FBuilder.Initialize(Mode := E_OrchestrationMode.ParallelSlots,
    TestCases := FCases);
AcceptedA := FBuilder.RegisterWithSlot(TestCase := ChildA,
    ExecutionSlot := 0);
Config := FBuilder.Finalize();
FZeroSlotRejectedMatches := NOT AcceptedA AND NOT Config.IsValid
    AND (FBuilder.Count = 0) AND (FCases[1] = 0)
    AND (FChildA.ExecutionSlot = CandidateSlotBeforeRejection);

FBuilder.Initialize(Mode := E_OrchestrationMode.ParallelSlots,
    TestCases := FCases);
AcceptedA := FBuilder.RegisterWithSlot(TestCase := ChildA,
    ExecutionSlot := 1);
AcceptedB := FBuilder.RegisterWithSlot(TestCase := ChildB,
    ExecutionSlot := 3);
Config := FBuilder.Finalize();
FSlotGapRejectedMatches := AcceptedA AND AcceptedB AND NOT Config.IsValid
    AND FBuilder.IsFinalized AND (FBuilder.Count = 2)
    AND (FCases[1] = ChildA) AND (FCases[2] = ChildB);
END_METHOD

END_FUNCTION_BLOCK

// ---- SelfTests/TestCases/TestSuite_TestSuiteConfigurationBuilder/Test_SuiteBuilderFinalizeReuse.TcPOU
{region 'Documentation'}
(*!
<summary>Checks empty and repeated finalization, sealed registration and a clean new build.</summary>
<description>Child mocks are inert interface identities and slot storage only; no child initialization or FB call is performed.</description>
*)
{endregion}
FUNCTION_BLOCK Test_SuiteBuilderFinalizeReuse EXTENDS TestCaseBase
VAR
    FBuilder : TestSuiteConfigurationBuilder;
    FCases : ARRAY[1..2] OF I_TestCase;
    FChildA : TestCaseMock;
    FChildB : TestCaseMock;
    FScenarioExecuted : BOOL;
    FChecksEvaluated : BOOL;
    FEmptyRejected : AssertTrue;
    FEmptyRejectedMatches : BOOL;
    FRepeatedFinalization : AssertTrue;
    FRepeatedFinalizationMatches : BOOL;
    FSealedRegistration : AssertTrue;
    FSealedRegistrationMatches : BOOL;
    FErrorRecorded : AssertTrue;
    FErrorRecordedMatches : BOOL;
    FFreshInitialize : AssertTrue;
    FFreshInitializeMatches : BOOL;
    FReuse : AssertTrue;
    FReuseMatches : BOOL;
END_VAR
VAR CONSTANT
    CandidateSlotBeforeRejection : UINT := 9;
END_VAR

SUPER^();

{region 'Documentation'}
(*!
<summary>Contributes each owned Assertion once without executing it.</summary>
*)
{endregion}
METHOD PROTECTED AggregateResults
VAR_INPUT
    Aggregator : I_ResultAggregator; //! Borrowed result sink owned by the outer Test Case; add this test's checking Assertions without resetting or retaining the sink.
END_VAR
Aggregator.AddProvider(Provider := FEmptyRejected);
Aggregator.AddProvider(Provider := FRepeatedFinalization);
Aggregator.AddProvider(Provider := FSealedRegistration);
Aggregator.AddProvider(Provider := FErrorRecorded);
Aggregator.AddProvider(Provider := FFreshInitialize);
Aggregator.AddProvider(Provider := FReuse);
END_METHOD

{region 'Documentation'}
(*!
<summary>Requires successful base and owned Assertion initialization.</summary>
*)
{endregion}
METHOD PROTECTED CheckInitialization : BOOL //! TRUE when the inherited initialization check and this concrete fixture check both accept the setup.
CheckInitialization := FALSE;
IF NOT SUPER^.CheckInitialization() THEN
    RETURN;
END_IF;

CheckInitialization := FEmptyRejected.IsInitialized
    AND FRepeatedFinalization.IsInitialized
    AND FSealedRegistration.IsInitialized
    AND FErrorRecorded.IsInitialized
    AND FFreshInitialize.IsInitialized
    AND FReuse.IsInitialized;
END_METHOD

{region 'Documentation'}
(*!
<summary>Configures one direct builder scenario and its named Assertions.</summary>
*)
{endregion}
METHOD PROTECTED Configure
FPreparationStateCount := 0;
FTestStateCount := 1;
FScenarioExecuted := FALSE;
FChecksEvaluated := FALSE;

FEmptyRejectedMatches := FALSE;
FEmptyRejected.Initialize(Parent := THIS^,
    AssertionName := 'EmptyRejected');
FRepeatedFinalizationMatches := FALSE;
FRepeatedFinalization.Initialize(Parent := THIS^,
    AssertionName := 'RepeatedFinalization');
FSealedRegistrationMatches := FALSE;
FSealedRegistration.Initialize(Parent := THIS^,
    AssertionName := 'SealedRegistration');
FErrorRecordedMatches := FALSE;
FErrorRecorded.Initialize(Parent := THIS^,
    AssertionName := 'ErrorRecorded');
FFreshInitializeMatches := FALSE;
FFreshInitialize.Initialize(Parent := THIS^,
    AssertionName := 'FreshInitialize');
FReuseMatches := FALSE;
FReuse.Initialize(Parent := THIS^,
    AssertionName := 'Reuse');
END_METHOD

{region 'Documentation'}
(*!
<summary>Completes Abort immediately; no asynchronous resource operation is started.</summary>
*)
{endregion}
METHOD PROTECTED ProcessAbort
VAR_INPUT
    Enable : BOOL; //! Phase permission supplied by the owning Test Case; FALSE does not authorize progression, while observation may continue.
END_VAR
IF Enable THEN
    CompleteAbort();
END_IF;
END_METHOD

{region 'Documentation'}
(*!
<summary>Evaluates recorded observations and consumes pending resets on disabled calls.</summary>
*)
{endregion}
METHOD PROTECTED ProcessAssertions
VAR_INPUT
    Enable : BOOL; //! Phase permission supplied by the owning Test Case; FALSE does not authorize progression, while observation may continue.
END_VAR
FEmptyRejected(Enable := Enable,
    State := State,
    IN := FEmptyRejectedMatches);

FRepeatedFinalization(Enable := Enable,
    State := State,
    IN := FRepeatedFinalizationMatches);

FSealedRegistration(Enable := Enable,
    State := State,
    IN := FSealedRegistrationMatches);

FErrorRecorded(Enable := Enable,
    State := State,
    IN := FErrorRecordedMatches);

FFreshInitialize(Enable := Enable,
    State := State,
    IN := FFreshInitializeMatches);

FReuse(Enable := Enable,
    State := State,
    IN := FReuseMatches);

IF Enable AND FEmptyRejected.EvaluationActive
    AND FRepeatedFinalization.EvaluationActive
    AND FSealedRegistration.EvaluationActive
    AND FErrorRecorded.EvaluationActive
    AND FFreshInitialize.EvaluationActive
    AND FReuse.EvaluationActive THEN
    FChecksEvaluated := TRUE;
END_IF;
END_METHOD

{region 'Documentation'}
(*!
<summary>No Preparation phase is needed for synchronous builder calls.</summary>
*)
{endregion}
METHOD PROTECTED ProcessPreparations
VAR_INPUT
    // SA0033: Required override signature; this scenario has no Preparation work.
    {attribute 'analysis' := '-33'}
    Enable : BOOL; //! Phase permission supplied by the owning Test Case; FALSE does not authorize progression, while observation may continue.
END_VAR
END_METHOD

{region 'Documentation'}
(*!
<summary>Clears recorded checks and Assertion results; each scenario initializes its own builder.</summary>
*)
{endregion}
METHOD PROTECTED ProcessReset
FScenarioExecuted := FALSE;
FChecksEvaluated := FALSE;
FEmptyRejectedMatches := FALSE;
FEmptyRejected.Reset();
FRepeatedFinalizationMatches := FALSE;
FRepeatedFinalization.Reset();
FSealedRegistrationMatches := FALSE;
FSealedRegistration.Reset();
FErrorRecordedMatches := FALSE;
FErrorRecorded.Reset();
FFreshInitializeMatches := FALSE;
FFreshInitialize.Reset();
FReuseMatches := FALSE;
FReuse.Reset();
CompleteReset();
END_METHOD

{region 'Documentation'}
(*!
<summary>Runs setup operations once, then completes after their observations have been evaluated.</summary>
*)
{endregion}
METHOD PROTECTED ProcessTests
VAR_INPUT
    Enable : BOOL; //! Phase permission supplied by the owning Test Case; FALSE does not authorize progression, while observation may continue.
END_VAR
IF NOT Enable THEN
    RETURN;
END_IF;

IF FChecksEvaluated THEN
    CompleteTests();
ELSIF NOT FScenarioExecuted THEN
    RunScenario();
    FScenarioExecuted := TRUE;
END_IF;
END_METHOD

{region 'Documentation'}
(*!
<summary>Checks empty and repeated finalization, sealed registration and a clean new build.</summary>
*)
{endregion}
METHOD PRIVATE RunScenario
VAR
    ChildA : I_TestCase;
    ChildB : I_TestCase;
    AcceptedA : BOOL;
    AcceptedB : BOOL;
    Config : ST_TestCaseCollectionConfig;
    RepeatedConfig : ST_TestCaseCollectionConfig;
END_VAR
ChildA := FChildA;
ChildB := FChildB;
FBuilder.Initialize(Mode := E_OrchestrationMode.Serial,
    TestCases := FCases);
Config := FBuilder.Finalize();
RepeatedConfig := FBuilder.Finalize();
FEmptyRejectedMatches := NOT Config.IsValid AND NOT RepeatedConfig.IsValid
    AND FBuilder.IsFinalized AND NOT FBuilder.IsValid AND (RepeatedConfig.Count = 0);

FBuilder.Initialize(Mode := E_OrchestrationMode.Serial,
    TestCases := FCases);
AcceptedA := FBuilder.Register(TestCase := ChildA);
Config := FBuilder.Finalize();
RepeatedConfig := FBuilder.Finalize();
FRepeatedFinalizationMatches := AcceptedA AND Config.IsValid AND RepeatedConfig.IsValid
    AND (RepeatedConfig.FirstIndex = Config.FirstIndex)
    AND (RepeatedConfig.LastIndex = Config.LastIndex)
    AND (RepeatedConfig.Count = Config.Count) AND (RepeatedConfig.Mode = Config.Mode);

FChildB.ExecutionSlot := CandidateSlotBeforeRejection;
AcceptedB := FBuilder.Register(TestCase := ChildB);
RepeatedConfig := FBuilder.Finalize();
FSealedRegistrationMatches := NOT AcceptedB AND RepeatedConfig.IsValid AND FBuilder.IsValid
    AND FBuilder.IsFinalized AND (FBuilder.Count = 1)
    AND (FCases[1] = ChildA) AND (FCases[2] = 0)
    AND (FChildB.ExecutionSlot = CandidateSlotBeforeRejection);

FBuilder.Initialize(Mode := E_OrchestrationMode.Serial,
    TestCases := FCases);
AcceptedA := FBuilder.Register(TestCase := ChildA);
AcceptedB := FBuilder.Register(TestCase := ChildA);
Config := FBuilder.Finalize();
FErrorRecordedMatches := AcceptedA AND NOT AcceptedB AND NOT Config.IsValid;

FBuilder.Initialize(Mode := E_OrchestrationMode.Parallel,
    TestCases := FCases);
FFreshInitializeMatches := NOT FBuilder.IsFinalized AND NOT FBuilder.IsValid
    AND (FBuilder.Count = 0) AND (FBuilder.Mode = E_OrchestrationMode.Parallel)
    AND (FCases[1] = 0) AND (FCases[2] = 0);
AcceptedB := FBuilder.Register(TestCase := ChildB);
Config := FBuilder.Finalize();
FReuseMatches := AcceptedB AND Config.IsValid AND FBuilder.IsValid AND FBuilder.IsFinalized
    AND (Config.Count = 1) AND (Config.Mode = E_OrchestrationMode.Parallel)
    AND (FCases[1] = ChildB) AND (FCases[2] = 0) AND (FChildB.ExecutionSlot = 1);
END_METHOD

END_FUNCTION_BLOCK

// ---- SelfTests/TestSuites/TestSuite_RunControlConfigurationBuilder.TcPOU
{region 'Documentation'}
(*!
<summary>Checks the Run Control builder directly without executing registered child lifecycles.</summary>
*)
{endregion}
FUNCTION_BLOCK TestSuite_RunControlConfigurationBuilder EXTENDS TestSuiteBase
VAR
    FSerial : Test_RunControlBuilderSerial;
    FParallel : Test_RunControlBuilderParallel;
    FSlotInsertion : Test_RunControlBuilderSlotInsertion;
    FCapacity : Test_RunControlBuilderCapacity;
    FRegistrationErrors : Test_RunControlBuilderRegistrationErrors;
    FFinalizeReuse : Test_RunControlBuilderFinalizeReuse;
    FTestCases : ARRAY[1..TestCaseCapacity] OF I_TestCase;
END_VAR
VAR CONSTANT
    TestCaseCapacity : UINT := 6;
END_VAR

SUPER^();

{region 'Documentation'}
(*!
<summary>Initializes and registers the six independent builder scenarios for serial execution.</summary>
*)
{endregion}
METHOD PROTECTED Configure
VAR_IN_OUT
    // SA0167: Borrowed owner builder; no temporary instance is created.
    {attribute 'analysis' := '-167'}
    Builder : TestSuiteConfigurationBuilder; //! Borrowed owner configuration builder used only during this Configure call; register this owner's concrete children.
END_VAR
VAR
    TestConfig : ST_TestCaseConfig;
END_VAR
Builder.Initialize(Mode := E_OrchestrationMode.Serial,
    TestCases := FTestCases);

FSerial.Initialize(Parent := THIS^,
    TestName := 'Serial',
    Config := TestConfig);
Builder.Register(TestCase := FSerial);

FParallel.Initialize(Parent := THIS^,
    TestName := 'Parallel',
    Config := TestConfig);
Builder.Register(TestCase := FParallel);

FSlotInsertion.Initialize(Parent := THIS^,
    TestName := 'SlotInsertion',
    Config := TestConfig);
Builder.Register(TestCase := FSlotInsertion);

FCapacity.Initialize(Parent := THIS^,
    TestName := 'Capacity',
    Config := TestConfig);
Builder.Register(TestCase := FCapacity);

FRegistrationErrors.Initialize(Parent := THIS^,
    TestName := 'RegistrationErrors',
    Config := TestConfig);
Builder.Register(TestCase := FRegistrationErrors);

FFinalizeReuse.Initialize(Parent := THIS^,
    TestName := 'FinalizeReuse',
    Config := TestConfig);
Builder.Register(TestCase := FFinalizeReuse);
END_METHOD

{region 'Documentation'}
(*!
<summary>Returns a registered scenario using the actual array index.</summary>
*)
{endregion}
METHOD PUBLIC GetTestCase : I_TestCase //! Typed child interface at the original array index; zero when no entry is available.
VAR_INPUT
    Index : DINT; //! Original occupied child-array index, rather than an ordinal position.
END_VAR
GetTestCase := 0;
IF (ChildCount = 0) OR (Index < ChildArrayLowerBound)
    OR (DINT_TO_LINT(Index) >= DINT_TO_LINT(ChildArrayLowerBound) + UINT_TO_LINT(ChildCount)) THEN
    RETURN;
END_IF;

GetTestCase := FTestCases[Index];
END_METHOD

{region 'Documentation'}
(*!
<summary>Calls the six owned scenarios once per initialized Suite cycle.</summary>
*)
{endregion}
METHOD PROTECTED ProcessTestCases
FSerial();
FParallel();
FSlotInsertion();
FCapacity();
FRegistrationErrors();
FFinalizeReuse();
END_METHOD

END_FUNCTION_BLOCK

// ---- SelfTests/TestCases/TestSuite_RunControlConfigurationBuilder/Test_RunControlBuilderSerial.TcPOU
{region 'Documentation'}
(*!
<summary>Checks Serial registration with shifted bounds and unused capacity.</summary>
<description>Child mocks are inert interface identities and slot storage only; no child initialization or FB call is performed.</description>
*)
{endregion}
FUNCTION_BLOCK Test_RunControlBuilderSerial EXTENDS TestCaseBase
VAR
    FBuilder : RunControlConfigurationBuilder;
    FSuites : ARRAY[4..7] OF I_TestSuite;
    FChildA : TestSuiteMock;
    FChildB : TestSuiteMock;
    FChildC : TestSuiteMock;
    FScenarioExecuted : BOOL;
    FChecksEvaluated : BOOL;
    FClearing : AssertTrue;
    FClearingMatches : BOOL;
    FRegistration : AssertTrue;
    FRegistrationMatches : BOOL;
    FOrder : AssertTrue;
    FOrderMatches : BOOL;
    FSlots : AssertTrue;
    FSlotsMatches : BOOL;
    FMetadata : AssertTrue;
    FMetadataMatches : BOOL;
    FFinalization : AssertTrue;
    FFinalizationMatches : BOOL;
END_VAR

SUPER^();

{region 'Documentation'}
(*!
<summary>Contributes each owned Assertion once without executing it.</summary>
*)
{endregion}
METHOD PROTECTED AggregateResults
VAR_INPUT
    Aggregator : I_ResultAggregator; //! Borrowed result sink owned by the outer Test Case; add this test's checking Assertions without resetting or retaining the sink.
END_VAR
Aggregator.AddProvider(Provider := FClearing);
Aggregator.AddProvider(Provider := FRegistration);
Aggregator.AddProvider(Provider := FOrder);
Aggregator.AddProvider(Provider := FSlots);
Aggregator.AddProvider(Provider := FMetadata);
Aggregator.AddProvider(Provider := FFinalization);
END_METHOD

{region 'Documentation'}
(*!
<summary>Requires successful base and owned Assertion initialization.</summary>
*)
{endregion}
METHOD PROTECTED CheckInitialization : BOOL //! TRUE when the inherited initialization check and this concrete fixture check both accept the setup.
CheckInitialization := FALSE;
IF NOT SUPER^.CheckInitialization() THEN
    RETURN;
END_IF;

CheckInitialization := FClearing.IsInitialized
    AND FRegistration.IsInitialized
    AND FOrder.IsInitialized
    AND FSlots.IsInitialized
    AND FMetadata.IsInitialized
    AND FFinalization.IsInitialized;
END_METHOD

{region 'Documentation'}
(*!
<summary>Configures one direct builder scenario and its named Assertions.</summary>
*)
{endregion}
METHOD PROTECTED Configure
FPreparationStateCount := 0;
FTestStateCount := 1;
FScenarioExecuted := FALSE;
FChecksEvaluated := FALSE;

FClearingMatches := FALSE;
FClearing.Initialize(Parent := THIS^,
    AssertionName := 'Clearing');
FRegistrationMatches := FALSE;
FRegistration.Initialize(Parent := THIS^,
    AssertionName := 'Registration');
FOrderMatches := FALSE;
FOrder.Initialize(Parent := THIS^,
    AssertionName := 'Order');
FSlotsMatches := FALSE;
FSlots.Initialize(Parent := THIS^,
    AssertionName := 'Slots');
FMetadataMatches := FALSE;
FMetadata.Initialize(Parent := THIS^,
    AssertionName := 'Metadata');
FFinalizationMatches := FALSE;
FFinalization.Initialize(Parent := THIS^,
    AssertionName := 'Finalization');
END_METHOD

{region 'Documentation'}
(*!
<summary>Completes Abort immediately; no asynchronous resource operation is started.</summary>
*)
{endregion}
METHOD PROTECTED ProcessAbort
VAR_INPUT
    Enable : BOOL; //! Phase permission supplied by the owning Test Case; FALSE does not authorize progression, while observation may continue.
END_VAR
IF Enable THEN
    CompleteAbort();
END_IF;
END_METHOD

{region 'Documentation'}
(*!
<summary>Evaluates recorded observations and consumes pending resets on disabled calls.</summary>
*)
{endregion}
METHOD PROTECTED ProcessAssertions
VAR_INPUT
    Enable : BOOL; //! Phase permission supplied by the owning Test Case; FALSE does not authorize progression, while observation may continue.
END_VAR
FClearing(Enable := Enable,
    State := State,
    IN := FClearingMatches);

FRegistration(Enable := Enable,
    State := State,
    IN := FRegistrationMatches);

FOrder(Enable := Enable,
    State := State,
    IN := FOrderMatches);

FSlots(Enable := Enable,
    State := State,
    IN := FSlotsMatches);

FMetadata(Enable := Enable,
    State := State,
    IN := FMetadataMatches);

FFinalization(Enable := Enable,
    State := State,
    IN := FFinalizationMatches);

IF Enable AND FClearing.EvaluationActive
    AND FRegistration.EvaluationActive
    AND FOrder.EvaluationActive
    AND FSlots.EvaluationActive
    AND FMetadata.EvaluationActive
    AND FFinalization.EvaluationActive THEN
    FChecksEvaluated := TRUE;
END_IF;
END_METHOD

{region 'Documentation'}
(*!
<summary>No Preparation phase is needed for synchronous builder calls.</summary>
*)
{endregion}
METHOD PROTECTED ProcessPreparations
VAR_INPUT
    // SA0033: Required override signature; this scenario has no Preparation work.
    {attribute 'analysis' := '-33'}
    Enable : BOOL; //! Phase permission supplied by the owning Test Case; FALSE does not authorize progression, while observation may continue.
END_VAR
END_METHOD

{region 'Documentation'}
(*!
<summary>Clears recorded checks and Assertion results; each scenario initializes its own builder.</summary>
*)
{endregion}
METHOD PROTECTED ProcessReset
FScenarioExecuted := FALSE;
FChecksEvaluated := FALSE;
FClearingMatches := FALSE;
FClearing.Reset();
FRegistrationMatches := FALSE;
FRegistration.Reset();
FOrderMatches := FALSE;
FOrder.Reset();
FSlotsMatches := FALSE;
FSlots.Reset();
FMetadataMatches := FALSE;
FMetadata.Reset();
FFinalizationMatches := FALSE;
FFinalization.Reset();
CompleteReset();
END_METHOD

{region 'Documentation'}
(*!
<summary>Runs setup operations once, then completes after their observations have been evaluated.</summary>
*)
{endregion}
METHOD PROTECTED ProcessTests
VAR_INPUT
    Enable : BOOL; //! Phase permission supplied by the owning Test Case; FALSE does not authorize progression, while observation may continue.
END_VAR
IF NOT Enable THEN
    RETURN;
END_IF;

IF FChecksEvaluated THEN
    CompleteTests();
ELSIF NOT FScenarioExecuted THEN
    RunScenario();
    FScenarioExecuted := TRUE;
END_IF;
END_METHOD

{region 'Documentation'}
(*!
<summary>Checks Serial registration with shifted bounds and unused capacity.</summary>
*)
{endregion}
METHOD PRIVATE RunScenario
VAR
    ChildA : I_TestSuite;
    ChildB : I_TestSuite;
    ChildC : I_TestSuite;
    AcceptedA : BOOL;
    AcceptedB : BOOL;
    AcceptedC : BOOL;
    Config : ST_TestSuiteCollectionConfig;
END_VAR
ChildA := FChildA;
ChildB := FChildB;
ChildC := FChildC;
FSuites[4] := ChildA;
FSuites[5] := ChildB;
FSuites[6] := ChildC;
FSuites[7] := ChildA;
FBuilder.Initialize(Mode := E_OrchestrationMode.Serial,
    TestSuites := FSuites);
FClearingMatches := (FSuites[4] = 0) AND (FSuites[5] = 0)
    AND (FSuites[6] = 0) AND (FSuites[7] = 0)
    AND (FBuilder.Count = 0) AND NOT FBuilder.IsValid AND NOT FBuilder.IsFinalized;

AcceptedA := FBuilder.Register(TestSuite := ChildC);
AcceptedB := FBuilder.Register(TestSuite := ChildA);
AcceptedC := FBuilder.Register(TestSuite := ChildB);
FRegistrationMatches := AcceptedA AND AcceptedB AND AcceptedC;
FOrderMatches := (FSuites[4] = ChildC) AND (FSuites[5] = ChildA)
    AND (FSuites[6] = ChildB) AND (FSuites[7] = 0);
FSlotsMatches := (FChildC.ExecutionSlot = 1) AND (FChildA.ExecutionSlot = 2)
    AND (FChildB.ExecutionSlot = 3);
FMetadataMatches := (FBuilder.FirstIndex = 4) AND (FBuilder.LastIndex = 7)
    AND (FBuilder.Count = 3) AND (FBuilder.Mode = E_OrchestrationMode.Serial);

Config := FBuilder.Finalize();
FFinalizationMatches := Config.IsValid AND FBuilder.IsValid AND FBuilder.IsFinalized
    AND (Config.FirstIndex = 4) AND (Config.LastIndex = 7) AND (Config.Count = 3)
    AND (Config.Mode = E_OrchestrationMode.Serial);
END_METHOD

END_FUNCTION_BLOCK

// ---- Framework/TestSuites/POU/TestSuiteMock.TcPOU
{region 'Documentation'}
(*!
<summary>Childless Suite double with simulated lifecycle, real owner events and real
reservations.</summary>
<description>
Initialize explicitly and let the parent reserve and dispatch Reset or Start. Call once per
task cycle. No Test Cases or Orchestrator are owned, and all child counters remain zero.

Ready gates Start; Completed and MinimumTestDuration gate normal completion. The minimum
defaults to T#100ms and survives Initialize and Reset. Error and Abort are not delayed.

Reset and Abort finish automatically without application acknowledgement. This mock validates
positive configured timeouts but does not reproduce child scheduling or child Reset/Abort
delays.
</description>
*)
{endregion}
FUNCTION_BLOCK TestSuiteMock IMPLEMENTS I_TestSuite
VAR_INPUT
    Ready : BOOL := TRUE; //! Application readiness gate for starting the mock; default TRUE.
    Completed : BOOL := TRUE; //! Allows normal mock completion after MinimumTestDuration; default TRUE.
    ResultValue : E_Result := E_Result.Passed; //! Simulated test outcome; default Passed. Lifecycle errors can still escalate the owner result.
END_VAR
VAR
    /// Instance binding; derived test adapters may assign it before first use.
    FEventPublisher : I_EventPublisher;
    FInitialized : BOOL;
    FConfigError : BOOL := TRUE;
    FName : STRING(GVL_Constants.NameLength);
    FResourceName : STRING(GVL_Constants.ResourceNameLength);
    FConfig : ST_TestSuiteConfig;
    FState : E_State := E_State.Uninitialized;
    FResult : E_Result := E_Result.NotEvaluated;
    FStatus : ST_TestSuiteStatus;
    FMethodRequests : ST_Command;
    FExecutionTimer : Stopwatch;
    FStateTimer : Stopwatch;
    FMinimumTestDuration : TIME := T#100ms;
    FExecutionSlot : UINT;
    FReservedEntryCount : UINT;
END_VAR
VAR_TEMP
    Requests : ST_Command;
END_VAR

ProcessRequests(InputRequests := FMethodRequests,
    Requests => Requests);
FExecutionTimer.Update();
FStateTimer.Update();
StateMachine(Requests := Requests);
UpdateStatus();
EmitFinalizationEvents();

{region 'Documentation'}
(*!
<summary>Publishes Result then Aggregation in the single Completing cycle, after result/status projection.</summary>
*)
{endregion}
METHOD PRIVATE EmitFinalizationEvents
IF FState <> E_State.Completing THEN
    RETURN;
END_IF;

PublishEvent(Event := CreateResultEvent(OwnerScope := E_OwnerScope.TestSuite,
    Name := FName,
    ResourceName := FResourceName,
    State := FState,
    Result := FResult,
    Message := ''));
PublishEvent(Event := CreateTestSuiteAggregationEvent(Name := FName,
    ResourceName := FResourceName,
    Status := FStatus));
END_METHOD

{region 'Documentation'}
(*!
<summary>Latches the technical Suite error and emits its first diagnostic; does not change state.</summary>
*)
{endregion}
METHOD PRIVATE Error
VAR_INPUT
    Message : STRING(GVL_Constants.MessageLength); //! Framework diagnostic text emitted only when first escalating the initialized, nonterminal mock result to Error.
END_VAR
IF (FState = E_State.Uninitialized) OR (FState = E_State.Completed) THEN
    RETURN;
END_IF;
IF FResult <> E_Result.Error THEN
    PublishEvent(Event := CreateFrameworkEvent(Name := FName,
        ResourceName := FResourceName,
        State := FState,
        Severity := E_EventSeverity.Error,
        Message := Message));
END_IF;
FResult := E_Result.Error;
END_METHOD

{region 'Documentation'}
(*!
<summary>Returns this instance's retained event-publication service.</summary>
<description>
If the local binding is zero, the getter takes GVL_EventBuffer.Publisher on access. An
established binding is retained; Initialize and lifecycle Reset do not replace it.

The default must be bound before first diagnostic use. Controlled test adapters may assign the
protected field before use. This getter performs no event publication, lifecycle processing or
reservation change.
</description>
*)
{endregion}
{attribute 'monitoring' := 'variable'}
PROPERTY PUBLIC EventPublisher : I_EventPublisher //! Returns this instance's retained event-publication service.
GET // PUBLIC
IF FEventPublisher = 0 THEN
    FEventPublisher := GVL_EventBuffer.Publisher;
END_IF;
EventPublisher := FEventPublisher;
END_GET
END_PROPERTY

{region 'Documentation'}
(*!
<summary>Parent-assigned configuration slot; Initialize and Reset retain it.</summary>
*)
{endregion}
{attribute 'monitoring' := 'call'}
PROPERTY PUBLIC ExecutionSlot : UINT //! Parent-assigned configuration slot; Initialize and Reset retain it.
GET // PUBLIC
ExecutionSlot := FExecutionSlot;
END_GET
SET // PUBLIC
FExecutionSlot := ExecutionSlot;
END_SET
END_PROPERTY

{region 'Documentation'}
(*!
<summary>Releases the own contribution only; this double has no children. Repeated release is
idempotent.</summary>
*)
{endregion}
METHOD PUBLIC FreeReservedEvents : BOOL //! TRUE when the own reservation is released or already zero; FALSE retains the unresolved contribution.
FreeReservedEvents := UpdateEventReservation(EntryCount := 0,
    HeadroomEntryCount := 0,
    ChildEntryCount := 0) = E_EventReservationResult.Accepted;
END_METHOD

{region 'Documentation'}
(*!
<summary>Reports configuration or runtime error.</summary>
*)
{endregion}
{attribute 'monitoring' := 'call'}
PROPERTY PUBLIC HasError : BOOL //! Reports configuration or runtime error.
GET // PUBLIC
HasError := FConfigError OR (FResult = E_Result.Error);
END_GET
END_PROPERTY

{region 'Documentation'}
(*!
<summary>Establishes the Suite identity and timing configuration without a child
collection.</summary>
<description>
Called by the parent at PLC startup; Reset preserves configuration and settings. Clears its
own old reservation after Event Buffer initialization; waits for the parent's Reset.

Reinitialization requires configuration reactivation or PLC Cold Reset followed by the
application's first-cycle initialization chain. Normal PLC Stop/Start and UnitTest Reset do not
rebuild configuration. Do not call Initialize as recovery during an active run.

The selected publisher must already be usable for configuration diagnostics. Failure leaves
IsInitialized FALSE; retained diagnostic identity is not proof of valid setup.
</description>
*)
{endregion}
METHOD PUBLIC Initialize : BOOL //! TRUE after successful identity and setup validation; FALSE leaves the object uninitialized.
VAR_INPUT
    Parent : I_RunControl; //! Owning Run Control with an established Name; read during Initialize, not retained.
    SuiteName : STRING(GVL_Constants.NameLength); //! Nonempty single name segment appended to Parent.Name; the complete name must fit NameLength.
    ResourceName : STRING(GVL_Constants.ResourceNameLength) := ''; //! Optional resource context for diagnostics; empty by default.
    Config : ST_TestSuiteConfig; //! Timeout configuration copied during initialization; all timeout values must be greater than zero.
END_VAR
VAR
    FullName : STRING(2 * GVL_Constants.NameLength + 1);
    EmptyStatus : ST_TestSuiteStatus;
END_VAR
Initialize := FALSE;
FInitialized := FALSE;
FReservedEntryCount := 0;
FConfigError := TRUE;
FState := E_State.Uninitialized;
FResult := E_Result.NotEvaluated;
FMethodRequests.Start := FALSE;
FMethodRequests.Abort := FALSE;
FMethodRequests.Reset := FALSE;
FExecutionTimer.Reset();
FStateTimer.Reset();
FStatus := EmptyStatus;
UpdateStatus();

FName := SuiteName;
FResourceName := ResourceName;
FConfig := Config;
IF Parent = 0 THEN
    PublishInitializationError(Message := 'Missing Run Control parent.');
    RETURN;
END_IF;
FullName := CONCAT(CONCAT(Parent.Name, '.'), SuiteName);
// SA0175: Bounded name projection; identity validation examines the full ASCII name.
{analysis -175}
FName := LEFT(FullName, UINT_TO_INT(GVL_Constants.NameLength));
{analysis +175}
IF NOT IsNameValid(Name := FullName, Depth := 2) THEN
    PublishInitializationError(Message := CONCAT('Invalid Test Suite name: ', FullName));
    RETURN;
END_IF;
IF (FConfig.Timeout = T#0ms) OR (FConfig.ResetTimeout = T#0ms) OR (FConfig.AbortTimeout = T#0ms) THEN
    PublishInitializationError(Message := 'Suite timeouts must be greater than zero.');
    RETURN;
END_IF;

FConfigError := FALSE;
FInitialized := TRUE;
UpdateStatus();
Initialize := TRUE;
END_METHOD

{region 'Documentation'}
(*!
<summary>Reports terminal completion, independently of the Completed input.</summary>
*)
{endregion}
{attribute 'monitoring' := 'call'}
PROPERTY PUBLIC IsComplete : BOOL //! Reports terminal completion, independently of the Completed input.
GET // PUBLIC
IsComplete := FState = E_State.Completed;
END_GET
END_PROPERTY

{region 'Documentation'}
(*!
<summary>Reports successful explicit identity and configuration initialization.</summary>
*)
{endregion}
{attribute 'monitoring' := 'call'}
PROPERTY PUBLIC IsInitialized : BOOL //! Reports successful explicit identity and configuration initialization.
GET // PUBLIC
IsInitialized := FInitialized;
END_GET
END_PROPERTY

{region 'Documentation'}
(*!
<summary>Start permission in initialized Idle, gated by the Ready input.</summary>
*)
{endregion}
{attribute 'monitoring' := 'call'}
PROPERTY PUBLIC IsReady : BOOL //! Start permission in initialized Idle, gated by the Ready input.
GET // PUBLIC
IsReady := FInitialized AND NOT FConfigError AND (FState = E_State.Idle)
    AND (FResult <> E_Result.Error) AND Ready;
END_GET
END_PROPERTY

{region 'Documentation'}
(*!
<summary>Minimum Running duration before normal completion; default T#100ms.</summary>
<description>
Zero permits immediate normal completion. Initialize and Reset retain this setting. Error,
explicit Abort and the configured execution timeout are not delayed.
</description>
*)
{endregion}
{attribute 'monitoring' := 'call'}
PROPERTY PUBLIC MinimumTestDuration : TIME //! Minimum Running duration before normal completion; default T#100ms.
GET // PUBLIC
MinimumTestDuration := FMinimumTestDuration;
END_GET
SET // PUBLIC
FMinimumTestDuration := MinimumTestDuration;
END_SET
END_PROPERTY

{region 'Documentation'}
(*!
<summary>Validated hierarchical Suite identity; rejected names may be retained truncated for
diagnosis.</summary>
*)
{endregion}
{attribute 'monitoring' := 'variable'}
PROPERTY PUBLIC Name : STRING(GVL_Constants.NameLength) //! Validated hierarchical Suite identity; rejected names may be retained truncated for diagnosis.
GET // PUBLIC
Name := FName;
END_GET
END_PROPERTY

{region 'Documentation'}
(*!
<summary>Consumes same-task requests, reports each received request and prioritizes Reset &gt; Abort &gt; Start.</summary>
<description>
Discards requests before initialization; never changes lifecycle state.
</description>
*)
{endregion}
METHOD PRIVATE ProcessRequests
VAR_IN_OUT
    InputRequests : ST_Command; //! Same-task request mailbox consumed and cleared, including before successful initialization.
END_VAR
VAR_OUTPUT
    Requests : ST_Command; //! Qualified request snapshot with Reset over Abort over Start; all FALSE before initialization.
END_VAR
Requests.Reset := FALSE;
Requests.Abort := FALSE;
Requests.Start := FALSE;

IF NOT FInitialized THEN
    InputRequests.Reset := FALSE;
    InputRequests.Abort := FALSE;
    InputRequests.Start := FALSE;
    RETURN;
END_IF;

Requests.Reset := InputRequests.Reset;
Requests.Abort := InputRequests.Abort AND NOT InputRequests.Reset;
Requests.Start := InputRequests.Start AND NOT InputRequests.Abort AND NOT InputRequests.Reset;

IF InputRequests.Reset THEN
    PublishEvent(Event := CreateResetEvent(OwnerScope := E_OwnerScope.TestSuite,
        Name := FName,
        ResourceName := FResourceName,
        State := FState));
END_IF;

IF InputRequests.Abort THEN
    PublishEvent(Event := CreateAbortEvent(OwnerScope := E_OwnerScope.TestSuite,
        Name := FName,
        ResourceName := FResourceName,
        State := FState));
END_IF;

IF InputRequests.Start THEN
    PublishEvent(Event := CreateStartEvent(OwnerScope := E_OwnerScope.TestSuite,
        Name := FName,
        ResourceName := FResourceName,
        State := FState));
END_IF;

InputRequests.Reset := FALSE;
InputRequests.Abort := FALSE;
InputRequests.Start := FALSE;
END_METHOD

{region 'Documentation'}
(*!
<summary>Publishes through the selected instance publisher without owning buffer loss accounting.</summary>
*)
{endregion}
METHOD PRIVATE PublishEvent
VAR_INPUT
    Event : ST_Event; //! Payload forwarded once through the selected usable publisher; no retry or local loss accounting.
END_VAR
EventPublisher.PublishEvent(Event := Event);
END_METHOD

{region 'Documentation'}
(*!
<summary>Emits a setup diagnostic without advancing lifecycle or changing the owner result.</summary>
*)
{endregion}
METHOD PRIVATE PublishInitializationError
VAR_INPUT
    Message : STRING(GVL_Constants.MessageLength); //! Setup diagnostic text sent through the required usable selected publisher without advancing lifecycle.
END_VAR
EventPublisher.PublishEvent(Event := CreateFrameworkEvent(Name := FName,
    ResourceName := FResourceName,
    State := E_State.Uninitialized,
    Severity := E_EventSeverity.Error,
    Message := Message));
END_METHOD

{region 'Documentation'}
(*!
<summary>Records an Abort request for the next regular FB call.</summary>
<description>
Repeated positive calls coalesce in the same-task request storage. Processing consumes the
requests with priority Reset, Abort, Start; calls before successful initialization are discarded
when processed.

Abort requests controlled termination of execution, not Reset cancellation. The owner
lifecycle determines whether the request applies.
</description>
*)
{endregion}
METHOD PUBLIC RequestAbort
FMethodRequests.Abort := TRUE;
END_METHOD

{region 'Documentation'}
(*!
<summary>Records a Reset request for the next regular FB call.</summary>
<description>
Repeated positive calls coalesce in the same-task request storage. Processing consumes the
requests with priority Reset, Abort, Start; calls before successful initialization are discarded
when processed.

Lifecycle Reset preserves configuration and publisher binding. It is not reinitialization or
Event Buffer Reset; capacity admission belongs to the parent when this object is a child.
</description>
*)
{endregion}
METHOD PUBLIC RequestReset
FMethodRequests.Reset := TRUE;
END_METHOD

{region 'Documentation'}
(*!
<summary>Records a Start request for the next regular FB call.</summary>
<description>
Repeated positive calls coalesce in the same-task request storage. Processing consumes the
requests with priority Reset, Abort, Start; calls before successful initialization are discarded
when processed.

Start is accepted by the lifecycle only in ready Idle. Recording the request does not start
execution synchronously.
</description>
*)
{endregion}
METHOD PUBLIC RequestStart
FMethodRequests.Start := TRUE;
END_METHOD

{region 'Documentation'}
(*!
<summary>Own contribution to the global Event Buffer reservation.</summary>
*)
{endregion}
{attribute 'monitoring' := 'call'}
PROPERTY PUBLIC ReservedEntryCount : UINT //! Own contribution to the global Event Buffer reservation.
GET // PUBLIC
ReservedEntryCount := FReservedEntryCount;
END_GET
END_PROPERTY

{region 'Documentation'}
(*!
<summary>Adjusts this owner's reservation to its execution budget immediately.</summary>
<description>
Only this owner's contribution is reserved; child budgets are separate. Local contribution and
publisher accounting are updated together without a lifecycle transition.

Accepted permits dispatch; WaitingForCapacity is retryable under the owner's timeout; Error
denotes invalid setup or an impossible budget. Calling before initialization reports a Framework
error. Repeated success aligns the total rather than adding a second budget.
</description>
*)
{endregion}
METHOD PUBLIC FINAL ReserveExecutionEvents : E_EventReservationResult //! Accepted on success, WaitingForCapacity for retryable pressure, Error for invalid setup or an impossible budget.
ReserveExecutionEvents := E_EventReservationResult.Error;
IF NOT FInitialized THEN
    PublishEvent(Event := CreateFrameworkEvent(Name := FName,
        ResourceName := FResourceName,
        State := FState,
        Severity := E_EventSeverity.Error,
        Message := 'ReserveExecutionEvents requires an initialized Test Suite.'));
    RETURN;
END_IF;

ReserveExecutionEvents := UpdateEventReservation(EntryCount := GVL_Constants.TestSuiteExecutionEventCount,
    HeadroomEntryCount := Param_EventBuffer.EventBufferExecutionHeadroom,
    ChildEntryCount := 0);
END_METHOD

{region 'Documentation'}
(*!
<summary>Adjusts this owner's reservation for capacity-admitted Reset immediately.</summary>
<description>
Does not dispatch Reset or clear existing events. Shared headroom and one Test Case Reset
allowance participate in admission, not this owner's stored contribution.

Accepted, WaitingForCapacity and Error distinguish success, temporary pressure and invalid
setup. An uninitialized call reports a Framework error. Lifecycle Reset must not silently clear the
reservation.

Although childless, the mock preserves the shared Suite admission rule with one unreserved Test Case Reset allowance. It reserves only its own Suite contribution and does not fabricate child reservations or events.
</description>
*)
{endregion}
METHOD PUBLIC FINAL ReserveResetEvents : E_EventReservationResult //! Accepted on success, WaitingForCapacity for retryable pressure, Error for invalid setup or an impossible budget.
ReserveResetEvents := E_EventReservationResult.Error;
IF NOT FInitialized THEN
    PublishEvent(Event := CreateFrameworkEvent(Name := FName,
        ResourceName := FResourceName,
        State := FState,
        Severity := E_EventSeverity.Error,
        Message := 'ReserveResetEvents requires an initialized Test Suite.'));
    RETURN;
END_IF;

ReserveResetEvents := UpdateEventReservation(EntryCount := GVL_Constants.TestSuiteResetEventCount,
    HeadroomEntryCount := Param_EventBuffer.EventBufferResetHeadroom,
    ChildEntryCount := GVL_Constants.TestCaseResetEventCount);
END_METHOD

{region 'Documentation'}
(*!
<summary>Held owner result; Reset clears it and Completed retains it.</summary>
*)
{endregion}
{attribute 'monitoring' := 'call'}
PROPERTY PUBLIC Result : E_Result //! Held owner result; Reset clears it and Completed retains it.
GET // PUBLIC
Result := FResult;
END_GET
END_PROPERTY

{region 'Documentation'}
(*!
<summary>Current simulated owner lifecycle state.</summary>
*)
{endregion}
{attribute 'monitoring' := 'call'}
PROPERTY PUBLIC State : E_State //! Current simulated owner lifecycle state.
GET // PUBLIC
State := FState;
END_GET
END_PROPERTY

{region 'Documentation'}
(*!
<summary>Processes simulated Suite transitions centrally; no child or Orchestrator execution.</summary>
<description>
Reset and Abort complete without external acknowledgement; Completed retains the result.

A new Reset request enters Reset without completing it in the same call. The next call enters Idle even if another Reset request is received; repeated requests during active Reset do not delay completion. Reset and Abort have no simulated delay or independent timeout supervision here; positive configured limits are validated at initialization, while execution Timeout is monitored. This double has no child scheduling.
</description>
*)
{endregion}
METHOD PRIVATE StateMachine
VAR_INPUT
    Requests : ST_Command; //! Consumed lifecycle request snapshot; a repeated Reset during active Reset permits the normal transition to Idle.
END_VAR
VAR
    PreviousState : E_State;
END_VAR
IF NOT FInitialized THEN
    RETURN;
END_IF;
PreviousState := FState;

IF Requests.Reset AND (FState <> E_State.Reset) THEN
    IF (FState = E_State.Starting) OR (FState = E_State.Running) OR (FState = E_State.Completing)
        OR (FState = E_State.Aborting) OR (FState = E_State.AbortingFromError) THEN
        PublishEvent(Event := CreateResetWarningEvent(OwnerScope := E_OwnerScope.TestSuite,
            Name := FName,
            ResourceName := FResourceName,
            State := FState));
    END_IF;
    FResult := E_Result.NotEvaluated;
    FExecutionTimer.Reset();
    FStateTimer.Reset();
    FState := E_State.Reset;
ELSE
    CASE FState OF
        E_State.Uninitialized:
            RETURN;

        E_State.Reset:
            FState := E_State.Idle;

        E_State.Idle:
            IF Requests.Start AND IsReady THEN
                FExecutionTimer.Start();
                FState := E_State.Starting;
            END_IF;

        E_State.Starting, E_State.Running:
            IF NOT FExecutionTimer.IsValid OR NOT FStateTimer.IsValid THEN
                Error(Message := 'Task clock error during Test Suite mock execution.');
            ELSIF FExecutionTimer.ElapsedLTime >= TIME_TO_LTIME(FConfig.Timeout) THEN
                Error(Message := 'Test Suite mock timeout reached.');
            ELSIF ResultValue = E_Result.Error THEN
                Error(Message := 'Test Suite mock reported an Error result.');
            ELSIF ResultValue = E_Result.Abort THEN
                Error(Message := 'Unexpected simulated result Abort; use RequestAbort.');
            END_IF;

            IF FResult = E_Result.Error THEN
                FExecutionTimer.Stop();
                FStateTimer.Stop();
                FState := E_State.AbortingFromError;
            ELSIF Requests.Abort THEN
                FResult := E_Result.Abort;
                FExecutionTimer.Stop();
                FStateTimer.Stop();
                FState := E_State.Aborting;
            ELSIF FState = E_State.Starting THEN
                FStateTimer.Start();
                FState := E_State.Running;
            ELSIF Completed AND (FStateTimer.ElapsedLTime >= TIME_TO_LTIME(FMinimumTestDuration)) THEN
                IF ResultValue = E_Result.Failed THEN
                    FResult := E_Result.Failed;
                ELSE
                    FResult := E_Result.Passed;
                END_IF;
                FExecutionTimer.Stop();
                FStateTimer.Stop();
                FState := E_State.Completing;
            END_IF;

        E_State.Completing:
            FState := E_State.Completed;

        E_State.Completed:
            RETURN;

        E_State.Aborting, E_State.AbortingFromError:
            IF (FState = E_State.Aborting) AND (ResultValue = E_Result.Error) THEN
                Error(Message := 'Test Suite mock reported an Error result during Abort.');
                FState := E_State.AbortingFromError;
            ELSE
                FState := E_State.Completing;
            END_IF;
    ELSE
        Error(Message := 'Unhandled Test Suite mock lifecycle state.');
        FExecutionTimer.Stop();
        FState := E_State.Completing;
    END_CASE;
END_IF;

IF FState <> PreviousState THEN
    PublishEvent(Event := CreateStateTransitionEvent(OwnerScope := E_OwnerScope.TestSuite,
        Name := FName,
        ResourceName := FResourceName,
        StateOld := PreviousState,
        StateNew := FState));
END_IF;
END_METHOD

{region 'Documentation'}
(*!
<summary>Current lifecycle and runtime snapshot; all Test Case counters are zero.</summary>
*)
{endregion}
PROPERTY PUBLIC Status : ST_TestSuiteStatus //! Current lifecycle and runtime snapshot; all Test Case counters are zero.
GET // PUBLIC
Status := FStatus;
END_GET
END_PROPERTY

{region 'Documentation'}
(*!
<summary>Checks own budget plus unreserved child allowance before changing either count.</summary>
<description>
Zero releases without capacity gating.

A zero target with no held contribution succeeds without publisher access. A nonzero held contribution is released through FreeReservedSpace without free-capacity gating. Positive targets check actual publisher validity/accounting and permanent capacity for target plus child allowance plus headroom. Temporary free capacity uses aggregate minus old own contribution plus target plus child allowance plus headroom. Even unchanged or reduced positive targets must pass this check. Only the Suite contribution changes; child allowance remains shared unreserved capacity. Failure leaves both ledgers unchanged.
</description>
*)
{endregion}
METHOD PRIVATE UpdateEventReservation : E_EventReservationResult //! Accepted after aligning the own contribution, WaitingForCapacity for temporary pressure, Error for invalid prerequisites or an impossible budget.
VAR_INPUT
    EntryCount : UINT; //! Target total own reservation, not an additional delta; zero releases the entire own contribution.
    HeadroomEntryCount : UINT; //! Shared unreserved producer headroom used in permanent and temporary capacity checks for positive targets.
    ChildEntryCount : UINT; //! Shared unreserved child allowance checked despite this mock having no concrete children; not stored as an own reservation.
END_VAR
VAR
    Publisher : I_EventPublisher;
    RequiredCapacity : UDINT;
    RequiredFreeEntries : UDINT;
END_VAR
UpdateEventReservation := E_EventReservationResult.Error;
IF (EntryCount = 0) AND (FReservedEntryCount = 0) THEN
    UpdateEventReservation := E_EventReservationResult.Accepted;
    RETURN;
END_IF;

Publisher := EventPublisher;

IF EntryCount = 0 THEN
    IF Publisher.FreeReservedSpace(EntryCount := FReservedEntryCount,
        OwnerReservedEntryCount := FReservedEntryCount) THEN
        UpdateEventReservation := E_EventReservationResult.Accepted;
    END_IF;
    RETURN;
END_IF;

IF NOT Publisher.IsValid THEN
    RETURN;
END_IF;
RequiredCapacity := UINT_TO_UDINT(EntryCount)
    + UINT_TO_UDINT(ChildEntryCount)
    + UINT_TO_UDINT(HeadroomEntryCount);
IF RequiredCapacity > UINT_TO_UDINT(Publisher.Capacity) THEN
    RETURN;
END_IF;
IF FReservedEntryCount > Publisher.ReservedEntryCount THEN
    RETURN;
END_IF;

RequiredFreeEntries := UINT_TO_UDINT(Publisher.ReservedEntryCount)
    - UINT_TO_UDINT(FReservedEntryCount)
    + UINT_TO_UDINT(EntryCount)
    + UINT_TO_UDINT(ChildEntryCount)
    + UINT_TO_UDINT(HeadroomEntryCount);
IF RequiredFreeEntries > UINT_TO_UDINT(Publisher.FreeEntryCount) THEN
    UpdateEventReservation := E_EventReservationResult.WaitingForCapacity;
    RETURN;
END_IF;

IF EntryCount < FReservedEntryCount THEN
    IF Publisher.FreeReservedSpace(EntryCount := FReservedEntryCount - EntryCount,
        OwnerReservedEntryCount := FReservedEntryCount) THEN
        UpdateEventReservation := E_EventReservationResult.Accepted;
    END_IF;
    RETURN;
END_IF;

IF Publisher.ReserveSpace(EntryCount := EntryCount - FReservedEntryCount,
    HeadroomEntryCount := HeadroomEntryCount,
    OwnerReservedEntryCount := FReservedEntryCount) THEN
    UpdateEventReservation := E_EventReservationResult.Accepted;
ELSE
    UpdateEventReservation := E_EventReservationResult.WaitingForCapacity;
END_IF;
END_METHOD

{region 'Documentation'}
(*!
<summary>Projects lifecycle and runtime each call; child counters remain zero because no children exist.</summary>
*)
{endregion}
METHOD PRIVATE UpdateStatus
VAR
    Execution : ST_ExecutionStatus;
END_VAR
Execution.State := FState;
Execution.Result := FResult;
Execution.ConfigError := FConfigError;
CASE FState OF
    E_State.Uninitialized:
        Execution.ExecutionStatus := E_ExecutionStatus.NotReady;
        Execution.Uninitialized := TRUE;
    E_State.Reset:
        Execution.ExecutionStatus := E_ExecutionStatus.Reset;
    E_State.Idle:
        Execution.ExecutionStatus := E_ExecutionStatus.Idle;
        Execution.Ready := IsReady;
    E_State.Starting:
        Execution.ExecutionStatus := E_ExecutionStatus.Starting;
    E_State.Running:
        Execution.ExecutionStatus := E_ExecutionStatus.Running;
        Execution.Running := TRUE;
    E_State.Completing:
        Execution.ExecutionStatus := E_ExecutionStatus.Completing;
    E_State.Completed:
        Execution.ExecutionStatus := E_ExecutionStatus.Completed;
        Execution.Completed := TRUE;
        Execution.Aborted := FResult = E_Result.Abort;
    E_State.Aborting, E_State.AbortingFromError:
        Execution.ExecutionStatus := E_ExecutionStatus.Aborting;
ELSE
    Execution.ExecutionStatus := E_ExecutionStatus.Error;
END_CASE;
Execution.Error := HasError;
FStatus.Execution := Execution;
FStatus.Runtime := FExecutionTimer.ElapsedTime;
END_METHOD

END_FUNCTION_BLOCK

// ---- SelfTests/TestCases/TestSuite_RunControlConfigurationBuilder/Test_RunControlBuilderParallel.TcPOU
{region 'Documentation'}
(*!
<summary>Checks Parallel registration order and shared slot across negative array bounds.</summary>
<description>Child mocks are inert interface identities and slot storage only; no child initialization or FB call is performed.</description>
*)
{endregion}
FUNCTION_BLOCK Test_RunControlBuilderParallel EXTENDS TestCaseBase
VAR
    FBuilder : RunControlConfigurationBuilder;
    FSuites : ARRAY[-2..1] OF I_TestSuite;
    FChildA : TestSuiteMock;
    FChildB : TestSuiteMock;
    FScenarioExecuted : BOOL;
    FChecksEvaluated : BOOL;
    FRegistration : AssertTrue;
    FRegistrationMatches : BOOL;
    FOrder : AssertTrue;
    FOrderMatches : BOOL;
    FSlots : AssertTrue;
    FSlotsMatches : BOOL;
    FMetadata : AssertTrue;
    FMetadataMatches : BOOL;
    FFinalization : AssertTrue;
    FFinalizationMatches : BOOL;
END_VAR

SUPER^();

{region 'Documentation'}
(*!
<summary>Contributes each owned Assertion once without executing it.</summary>
*)
{endregion}
METHOD PROTECTED AggregateResults
VAR_INPUT
    Aggregator : I_ResultAggregator; //! Borrowed result sink owned by the outer Test Case; add this test's checking Assertions without resetting or retaining the sink.
END_VAR
Aggregator.AddProvider(Provider := FRegistration);
Aggregator.AddProvider(Provider := FOrder);
Aggregator.AddProvider(Provider := FSlots);
Aggregator.AddProvider(Provider := FMetadata);
Aggregator.AddProvider(Provider := FFinalization);
END_METHOD

{region 'Documentation'}
(*!
<summary>Requires successful base and owned Assertion initialization.</summary>
*)
{endregion}
METHOD PROTECTED CheckInitialization : BOOL //! TRUE when the inherited initialization check and this concrete fixture check both accept the setup.
CheckInitialization := FALSE;
IF NOT SUPER^.CheckInitialization() THEN
    RETURN;
END_IF;

CheckInitialization := FRegistration.IsInitialized
    AND FOrder.IsInitialized
    AND FSlots.IsInitialized
    AND FMetadata.IsInitialized
    AND FFinalization.IsInitialized;
END_METHOD

{region 'Documentation'}
(*!
<summary>Configures one direct builder scenario and its named Assertions.</summary>
*)
{endregion}
METHOD PROTECTED Configure
FPreparationStateCount := 0;
FTestStateCount := 1;
FScenarioExecuted := FALSE;
FChecksEvaluated := FALSE;

FRegistrationMatches := FALSE;
FRegistration.Initialize(Parent := THIS^,
    AssertionName := 'Registration');
FOrderMatches := FALSE;
FOrder.Initialize(Parent := THIS^,
    AssertionName := 'Order');
FSlotsMatches := FALSE;
FSlots.Initialize(Parent := THIS^,
    AssertionName := 'Slots');
FMetadataMatches := FALSE;
FMetadata.Initialize(Parent := THIS^,
    AssertionName := 'Metadata');
FFinalizationMatches := FALSE;
FFinalization.Initialize(Parent := THIS^,
    AssertionName := 'Finalization');
END_METHOD

{region 'Documentation'}
(*!
<summary>Completes Abort immediately; no asynchronous resource operation is started.</summary>
*)
{endregion}
METHOD PROTECTED ProcessAbort
VAR_INPUT
    Enable : BOOL; //! Phase permission supplied by the owning Test Case; FALSE does not authorize progression, while observation may continue.
END_VAR
IF Enable THEN
    CompleteAbort();
END_IF;
END_METHOD

{region 'Documentation'}
(*!
<summary>Evaluates recorded observations and consumes pending resets on disabled calls.</summary>
*)
{endregion}
METHOD PROTECTED ProcessAssertions
VAR_INPUT
    Enable : BOOL; //! Phase permission supplied by the owning Test Case; FALSE does not authorize progression, while observation may continue.
END_VAR
FRegistration(Enable := Enable,
    State := State,
    IN := FRegistrationMatches);

FOrder(Enable := Enable,
    State := State,
    IN := FOrderMatches);

FSlots(Enable := Enable,
    State := State,
    IN := FSlotsMatches);

FMetadata(Enable := Enable,
    State := State,
    IN := FMetadataMatches);

FFinalization(Enable := Enable,
    State := State,
    IN := FFinalizationMatches);

IF Enable AND FRegistration.EvaluationActive
    AND FOrder.EvaluationActive
    AND FSlots.EvaluationActive
    AND FMetadata.EvaluationActive
    AND FFinalization.EvaluationActive THEN
    FChecksEvaluated := TRUE;
END_IF;
END_METHOD

{region 'Documentation'}
(*!
<summary>No Preparation phase is needed for synchronous builder calls.</summary>
*)
{endregion}
METHOD PROTECTED ProcessPreparations
VAR_INPUT
    // SA0033: Required override signature; this scenario has no Preparation work.
    {attribute 'analysis' := '-33'}
    Enable : BOOL; //! Phase permission supplied by the owning Test Case; FALSE does not authorize progression, while observation may continue.
END_VAR
END_METHOD

{region 'Documentation'}
(*!
<summary>Clears recorded checks and Assertion results; each scenario initializes its own builder.</summary>
*)
{endregion}
METHOD PROTECTED ProcessReset
FScenarioExecuted := FALSE;
FChecksEvaluated := FALSE;
FRegistrationMatches := FALSE;
FRegistration.Reset();
FOrderMatches := FALSE;
FOrder.Reset();
FSlotsMatches := FALSE;
FSlots.Reset();
FMetadataMatches := FALSE;
FMetadata.Reset();
FFinalizationMatches := FALSE;
FFinalization.Reset();
CompleteReset();
END_METHOD

{region 'Documentation'}
(*!
<summary>Runs setup operations once, then completes after their observations have been evaluated.</summary>
*)
{endregion}
METHOD PROTECTED ProcessTests
VAR_INPUT
    Enable : BOOL; //! Phase permission supplied by the owning Test Case; FALSE does not authorize progression, while observation may continue.
END_VAR
IF NOT Enable THEN
    RETURN;
END_IF;

IF FChecksEvaluated THEN
    CompleteTests();
ELSIF NOT FScenarioExecuted THEN
    RunScenario();
    FScenarioExecuted := TRUE;
END_IF;
END_METHOD

{region 'Documentation'}
(*!
<summary>Checks Parallel registration order and shared slot across negative array bounds.</summary>
*)
{endregion}
METHOD PRIVATE RunScenario
VAR
    ChildA : I_TestSuite;
    ChildB : I_TestSuite;
    AcceptedA : BOOL;
    AcceptedB : BOOL;
    Config : ST_TestSuiteCollectionConfig;
END_VAR
ChildA := FChildA;
ChildB := FChildB;
FBuilder.Initialize(Mode := E_OrchestrationMode.Parallel,
    TestSuites := FSuites);
AcceptedA := FBuilder.Register(TestSuite := ChildB);
AcceptedB := FBuilder.Register(TestSuite := ChildA);
FRegistrationMatches := AcceptedA AND AcceptedB;
FOrderMatches := (FSuites[-2] = ChildB) AND (FSuites[-1] = ChildA)
    AND (FSuites[0] = 0) AND (FSuites[1] = 0);
FSlotsMatches := (FChildA.ExecutionSlot = 1) AND (FChildB.ExecutionSlot = 1);
FMetadataMatches := (FBuilder.FirstIndex = -2) AND (FBuilder.LastIndex = 1)
    AND (FBuilder.Count = 2) AND (FBuilder.Mode = E_OrchestrationMode.Parallel);

Config := FBuilder.Finalize();
FFinalizationMatches := Config.IsValid AND FBuilder.IsValid AND FBuilder.IsFinalized
    AND (Config.FirstIndex = -2) AND (Config.LastIndex = 1) AND (Config.Count = 2)
    AND (Config.Mode = E_OrchestrationMode.Parallel);
END_METHOD

END_FUNCTION_BLOCK

// ---- SelfTests/TestCases/TestSuite_RunControlConfigurationBuilder/Test_RunControlBuilderSlotInsertion.TcPOU
{region 'Documentation'}
(*!
<summary>Checks stable insertion into two slots, including a temporary gap before Finalize.</summary>
<description>Child mocks are inert interface identities and slot storage only; no child initialization or FB call is performed.</description>
*)
{endregion}
FUNCTION_BLOCK Test_RunControlBuilderSlotInsertion EXTENDS TestCaseBase
VAR
    FBuilder : RunControlConfigurationBuilder;
    FSuites : ARRAY[1..4] OF I_TestSuite;
    FChildA : TestSuiteMock;
    FChildB : TestSuiteMock;
    FChildC : TestSuiteMock;
    FChildD : TestSuiteMock;
    FScenarioExecuted : BOOL;
    FChecksEvaluated : BOOL;
    FRegistration : AssertTrue;
    FRegistrationMatches : BOOL;
    FOrder : AssertTrue;
    FOrderMatches : BOOL;
    FSlots : AssertTrue;
    FSlotsMatches : BOOL;
    FFinalization : AssertTrue;
    FFinalizationMatches : BOOL;
END_VAR

SUPER^();

{region 'Documentation'}
(*!
<summary>Contributes each owned Assertion once without executing it.</summary>
*)
{endregion}
METHOD PROTECTED AggregateResults
VAR_INPUT
    Aggregator : I_ResultAggregator; //! Borrowed result sink owned by the outer Test Case; add this test's checking Assertions without resetting or retaining the sink.
END_VAR
Aggregator.AddProvider(Provider := FRegistration);
Aggregator.AddProvider(Provider := FOrder);
Aggregator.AddProvider(Provider := FSlots);
Aggregator.AddProvider(Provider := FFinalization);
END_METHOD

{region 'Documentation'}
(*!
<summary>Requires successful base and owned Assertion initialization.</summary>
*)
{endregion}
METHOD PROTECTED CheckInitialization : BOOL //! TRUE when the inherited initialization check and this concrete fixture check both accept the setup.
CheckInitialization := FALSE;
IF NOT SUPER^.CheckInitialization() THEN
    RETURN;
END_IF;

CheckInitialization := FRegistration.IsInitialized
    AND FOrder.IsInitialized
    AND FSlots.IsInitialized
    AND FFinalization.IsInitialized;
END_METHOD

{region 'Documentation'}
(*!
<summary>Configures one direct builder scenario and its named Assertions.</summary>
*)
{endregion}
METHOD PROTECTED Configure
FPreparationStateCount := 0;
FTestStateCount := 1;
FScenarioExecuted := FALSE;
FChecksEvaluated := FALSE;

FRegistrationMatches := FALSE;
FRegistration.Initialize(Parent := THIS^,
    AssertionName := 'Registration');
FOrderMatches := FALSE;
FOrder.Initialize(Parent := THIS^,
    AssertionName := 'Order');
FSlotsMatches := FALSE;
FSlots.Initialize(Parent := THIS^,
    AssertionName := 'Slots');
FFinalizationMatches := FALSE;
FFinalization.Initialize(Parent := THIS^,
    AssertionName := 'Finalization');
END_METHOD

{region 'Documentation'}
(*!
<summary>Completes Abort immediately; no asynchronous resource operation is started.</summary>
*)
{endregion}
METHOD PROTECTED ProcessAbort
VAR_INPUT
    Enable : BOOL; //! Phase permission supplied by the owning Test Case; FALSE does not authorize progression, while observation may continue.
END_VAR
IF Enable THEN
    CompleteAbort();
END_IF;
END_METHOD

{region 'Documentation'}
(*!
<summary>Evaluates recorded observations and consumes pending resets on disabled calls.</summary>
*)
{endregion}
METHOD PROTECTED ProcessAssertions
VAR_INPUT
    Enable : BOOL; //! Phase permission supplied by the owning Test Case; FALSE does not authorize progression, while observation may continue.
END_VAR
FRegistration(Enable := Enable,
    State := State,
    IN := FRegistrationMatches);

FOrder(Enable := Enable,
    State := State,
    IN := FOrderMatches);

FSlots(Enable := Enable,
    State := State,
    IN := FSlotsMatches);

FFinalization(Enable := Enable,
    State := State,
    IN := FFinalizationMatches);

IF Enable AND FRegistration.EvaluationActive
    AND FOrder.EvaluationActive
    AND FSlots.EvaluationActive
    AND FFinalization.EvaluationActive THEN
    FChecksEvaluated := TRUE;
END_IF;
END_METHOD

{region 'Documentation'}
(*!
<summary>No Preparation phase is needed for synchronous builder calls.</summary>
*)
{endregion}
METHOD PROTECTED ProcessPreparations
VAR_INPUT
    // SA0033: Required override signature; this scenario has no Preparation work.
    {attribute 'analysis' := '-33'}
    Enable : BOOL; //! Phase permission supplied by the owning Test Case; FALSE does not authorize progression, while observation may continue.
END_VAR
END_METHOD

{region 'Documentation'}
(*!
<summary>Clears recorded checks and Assertion results; each scenario initializes its own builder.</summary>
*)
{endregion}
METHOD PROTECTED ProcessReset
FScenarioExecuted := FALSE;
FChecksEvaluated := FALSE;
FRegistrationMatches := FALSE;
FRegistration.Reset();
FOrderMatches := FALSE;
FOrder.Reset();
FSlotsMatches := FALSE;
FSlots.Reset();
FFinalizationMatches := FALSE;
FFinalization.Reset();
CompleteReset();
END_METHOD

{region 'Documentation'}
(*!
<summary>Runs setup operations once, then completes after their observations have been evaluated.</summary>
*)
{endregion}
METHOD PROTECTED ProcessTests
VAR_INPUT
    Enable : BOOL; //! Phase permission supplied by the owning Test Case; FALSE does not authorize progression, while observation may continue.
END_VAR
IF NOT Enable THEN
    RETURN;
END_IF;

IF FChecksEvaluated THEN
    CompleteTests();
ELSIF NOT FScenarioExecuted THEN
    RunScenario();
    FScenarioExecuted := TRUE;
END_IF;
END_METHOD

{region 'Documentation'}
(*!
<summary>Checks stable insertion into two slots, including a temporary gap before Finalize.</summary>
*)
{endregion}
METHOD PRIVATE RunScenario
VAR
    ChildA : I_TestSuite;
    ChildB : I_TestSuite;
    ChildC : I_TestSuite;
    ChildD : I_TestSuite;
    AcceptedA : BOOL;
    AcceptedB : BOOL;
    AcceptedC : BOOL;
    AcceptedD : BOOL;
    Config : ST_TestSuiteCollectionConfig;
END_VAR
ChildA := FChildA;
ChildB := FChildB;
ChildC := FChildC;
ChildD := FChildD;
FBuilder.Initialize(Mode := E_OrchestrationMode.ParallelSlots,
    TestSuites := FSuites);
AcceptedA := FBuilder.RegisterWithSlot(TestSuite := ChildA,
    ExecutionSlot := 2);
AcceptedB := FBuilder.RegisterWithSlot(TestSuite := ChildB,
    ExecutionSlot := 1);
AcceptedC := FBuilder.RegisterWithSlot(TestSuite := ChildC,
    ExecutionSlot := 2);
AcceptedD := FBuilder.RegisterWithSlot(TestSuite := ChildD,
    ExecutionSlot := 1);
FRegistrationMatches := AcceptedA AND AcceptedB AND AcceptedC AND AcceptedD;
FOrderMatches := (FSuites[1] = ChildB) AND (FSuites[2] = ChildD)
    AND (FSuites[3] = ChildA) AND (FSuites[4] = ChildC);
FSlotsMatches := (FChildA.ExecutionSlot = 2) AND (FChildB.ExecutionSlot = 1)
    AND (FChildC.ExecutionSlot = 2) AND (FChildD.ExecutionSlot = 1);

Config := FBuilder.Finalize();
FFinalizationMatches := Config.IsValid AND FBuilder.IsValid AND FBuilder.IsFinalized
    AND (Config.FirstIndex = 1) AND (Config.LastIndex = 4) AND (Config.Count = 4)
    AND (Config.Mode = E_OrchestrationMode.ParallelSlots);
END_METHOD

END_FUNCTION_BLOCK

// ---- SelfTests/TestCases/TestSuite_RunControlConfigurationBuilder/Test_RunControlBuilderCapacity.TcPOU
{region 'Documentation'}
(*!
<summary>Checks exact capacity and rejection before array or candidate-slot mutation.</summary>
<description>Child mocks are inert interface identities and slot storage only; no child initialization or FB call is performed.</description>
*)
{endregion}
FUNCTION_BLOCK Test_RunControlBuilderCapacity EXTENDS TestCaseBase
VAR
    FBuilder : RunControlConfigurationBuilder;
    FSuites : ARRAY[1..2] OF I_TestSuite;
    FChildA : TestSuiteMock;
    FChildB : TestSuiteMock;
    FChildC : TestSuiteMock;
    FScenarioExecuted : BOOL;
    FChecksEvaluated : BOOL;
    FExactCapacity : AssertTrue;
    FExactCapacityMatches : BOOL;
    FOverflowRejected : AssertTrue;
    FOverflowRejectedMatches : BOOL;
    FCompositionPreserved : AssertTrue;
    FCompositionPreservedMatches : BOOL;
    FErrorLatched : AssertTrue;
    FErrorLatchedMatches : BOOL;
END_VAR
VAR CONSTANT
    CandidateSlotBeforeRejection : UINT := 9;
END_VAR

SUPER^();

{region 'Documentation'}
(*!
<summary>Contributes each owned Assertion once without executing it.</summary>
*)
{endregion}
METHOD PROTECTED AggregateResults
VAR_INPUT
    Aggregator : I_ResultAggregator; //! Borrowed result sink owned by the outer Test Case; add this test's checking Assertions without resetting or retaining the sink.
END_VAR
Aggregator.AddProvider(Provider := FExactCapacity);
Aggregator.AddProvider(Provider := FOverflowRejected);
Aggregator.AddProvider(Provider := FCompositionPreserved);
Aggregator.AddProvider(Provider := FErrorLatched);
END_METHOD

{region 'Documentation'}
(*!
<summary>Requires successful base and owned Assertion initialization.</summary>
*)
{endregion}
METHOD PROTECTED CheckInitialization : BOOL //! TRUE when the inherited initialization check and this concrete fixture check both accept the setup.
CheckInitialization := FALSE;
IF NOT SUPER^.CheckInitialization() THEN
    RETURN;
END_IF;

CheckInitialization := FExactCapacity.IsInitialized
    AND FOverflowRejected.IsInitialized
    AND FCompositionPreserved.IsInitialized
    AND FErrorLatched.IsInitialized;
END_METHOD

{region 'Documentation'}
(*!
<summary>Configures one direct builder scenario and its named Assertions.</summary>
*)
{endregion}
METHOD PROTECTED Configure
FPreparationStateCount := 0;
FTestStateCount := 1;
FScenarioExecuted := FALSE;
FChecksEvaluated := FALSE;

FExactCapacityMatches := FALSE;
FExactCapacity.Initialize(Parent := THIS^,
    AssertionName := 'ExactCapacity');
FOverflowRejectedMatches := FALSE;
FOverflowRejected.Initialize(Parent := THIS^,
    AssertionName := 'OverflowRejected');
FCompositionPreservedMatches := FALSE;
FCompositionPreserved.Initialize(Parent := THIS^,
    AssertionName := 'CompositionPreserved');
FErrorLatchedMatches := FALSE;
FErrorLatched.Initialize(Parent := THIS^,
    AssertionName := 'ErrorLatched');
END_METHOD

{region 'Documentation'}
(*!
<summary>Completes Abort immediately; no asynchronous resource operation is started.</summary>
*)
{endregion}
METHOD PROTECTED ProcessAbort
VAR_INPUT
    Enable : BOOL; //! Phase permission supplied by the owning Test Case; FALSE does not authorize progression, while observation may continue.
END_VAR
IF Enable THEN
    CompleteAbort();
END_IF;
END_METHOD

{region 'Documentation'}
(*!
<summary>Evaluates recorded observations and consumes pending resets on disabled calls.</summary>
*)
{endregion}
METHOD PROTECTED ProcessAssertions
VAR_INPUT
    Enable : BOOL; //! Phase permission supplied by the owning Test Case; FALSE does not authorize progression, while observation may continue.
END_VAR
FExactCapacity(Enable := Enable,
    State := State,
    IN := FExactCapacityMatches);

FOverflowRejected(Enable := Enable,
    State := State,
    IN := FOverflowRejectedMatches);

FCompositionPreserved(Enable := Enable,
    State := State,
    IN := FCompositionPreservedMatches);

FErrorLatched(Enable := Enable,
    State := State,
    IN := FErrorLatchedMatches);

IF Enable AND FExactCapacity.EvaluationActive
    AND FOverflowRejected.EvaluationActive
    AND FCompositionPreserved.EvaluationActive
    AND FErrorLatched.EvaluationActive THEN
    FChecksEvaluated := TRUE;
END_IF;
END_METHOD

{region 'Documentation'}
(*!
<summary>No Preparation phase is needed for synchronous builder calls.</summary>
*)
{endregion}
METHOD PROTECTED ProcessPreparations
VAR_INPUT
    // SA0033: Required override signature; this scenario has no Preparation work.
    {attribute 'analysis' := '-33'}
    Enable : BOOL; //! Phase permission supplied by the owning Test Case; FALSE does not authorize progression, while observation may continue.
END_VAR
END_METHOD

{region 'Documentation'}
(*!
<summary>Clears recorded checks and Assertion results; each scenario initializes its own builder.</summary>
*)
{endregion}
METHOD PROTECTED ProcessReset
FScenarioExecuted := FALSE;
FChecksEvaluated := FALSE;
FExactCapacityMatches := FALSE;
FExactCapacity.Reset();
FOverflowRejectedMatches := FALSE;
FOverflowRejected.Reset();
FCompositionPreservedMatches := FALSE;
FCompositionPreserved.Reset();
FErrorLatchedMatches := FALSE;
FErrorLatched.Reset();
CompleteReset();
END_METHOD

{region 'Documentation'}
(*!
<summary>Runs setup operations once, then completes after their observations have been evaluated.</summary>
*)
{endregion}
METHOD PROTECTED ProcessTests
VAR_INPUT
    Enable : BOOL; //! Phase permission supplied by the owning Test Case; FALSE does not authorize progression, while observation may continue.
END_VAR
IF NOT Enable THEN
    RETURN;
END_IF;

IF FChecksEvaluated THEN
    CompleteTests();
ELSIF NOT FScenarioExecuted THEN
    RunScenario();
    FScenarioExecuted := TRUE;
END_IF;
END_METHOD

{region 'Documentation'}
(*!
<summary>Checks exact capacity and rejection before array or candidate-slot mutation.</summary>
*)
{endregion}
METHOD PRIVATE RunScenario
VAR
    ChildA : I_TestSuite;
    ChildB : I_TestSuite;
    ChildC : I_TestSuite;
    AcceptedA : BOOL;
    AcceptedB : BOOL;
    AcceptedC : BOOL;
    Config : ST_TestSuiteCollectionConfig;
END_VAR
ChildA := FChildA;
ChildB := FChildB;
ChildC := FChildC;
FBuilder.Initialize(Mode := E_OrchestrationMode.Serial,
    TestSuites := FSuites);
AcceptedA := FBuilder.Register(TestSuite := ChildA);
AcceptedB := FBuilder.Register(TestSuite := ChildB);
Config := FBuilder.Finalize();
FExactCapacityMatches := AcceptedA AND AcceptedB AND Config.IsValid
    AND (Config.Count = 2) AND (FSuites[1] = ChildA) AND (FSuites[2] = ChildB);

FBuilder.Initialize(Mode := E_OrchestrationMode.Serial,
    TestSuites := FSuites);
AcceptedA := FBuilder.Register(TestSuite := ChildA);
AcceptedB := FBuilder.Register(TestSuite := ChildB);
FChildC.ExecutionSlot := CandidateSlotBeforeRejection;
AcceptedC := FBuilder.Register(TestSuite := ChildC);
FOverflowRejectedMatches := AcceptedA AND AcceptedB AND NOT AcceptedC;
FCompositionPreservedMatches := (FBuilder.Count = 2)
    AND (FSuites[1] = ChildA) AND (FSuites[2] = ChildB)
    AND (FChildA.ExecutionSlot = 1) AND (FChildB.ExecutionSlot = 2)
    AND (FChildC.ExecutionSlot = CandidateSlotBeforeRejection);

Config := FBuilder.Finalize();
FErrorLatchedMatches := NOT Config.IsValid AND NOT FBuilder.IsValid
    AND FBuilder.IsFinalized AND (Config.Count = 2);
END_METHOD

END_FUNCTION_BLOCK

// ---- SelfTests/TestCases/TestSuite_RunControlConfigurationBuilder/Test_RunControlBuilderRegistrationErrors.TcPOU
{region 'Documentation'}
(*!
<summary>Checks typical setup mistakes without executing the registered child objects.</summary>
<description>Child mocks are inert interface identities and slot storage only; no child initialization or FB call is performed.</description>
*)
{endregion}
FUNCTION_BLOCK Test_RunControlBuilderRegistrationErrors EXTENDS TestCaseBase
VAR
    FBuilder : RunControlConfigurationBuilder;
    FSuites : ARRAY[1..2] OF I_TestSuite;
    FChildA : TestSuiteMock;
    FChildB : TestSuiteMock;
    FScenarioExecuted : BOOL;
    FChecksEvaluated : BOOL;
    FDuplicateRejected : AssertTrue;
    FDuplicateRejectedMatches : BOOL;
    FNullRejected : AssertTrue;
    FNullRejectedMatches : BOOL;
    FExplicitSlotRejected : AssertTrue;
    FExplicitSlotRejectedMatches : BOOL;
    FMissingSlotRejected : AssertTrue;
    FMissingSlotRejectedMatches : BOOL;
    FZeroSlotRejected : AssertTrue;
    FZeroSlotRejectedMatches : BOOL;
    FSlotGapRejected : AssertTrue;
    FSlotGapRejectedMatches : BOOL;
END_VAR
VAR CONSTANT
    CandidateSlotBeforeRejection : UINT := 9;
END_VAR

SUPER^();

{region 'Documentation'}
(*!
<summary>Contributes each owned Assertion once without executing it.</summary>
*)
{endregion}
METHOD PROTECTED AggregateResults
VAR_INPUT
    Aggregator : I_ResultAggregator; //! Borrowed result sink owned by the outer Test Case; add this test's checking Assertions without resetting or retaining the sink.
END_VAR
Aggregator.AddProvider(Provider := FDuplicateRejected);
Aggregator.AddProvider(Provider := FNullRejected);
Aggregator.AddProvider(Provider := FExplicitSlotRejected);
Aggregator.AddProvider(Provider := FMissingSlotRejected);
Aggregator.AddProvider(Provider := FZeroSlotRejected);
Aggregator.AddProvider(Provider := FSlotGapRejected);
END_METHOD

{region 'Documentation'}
(*!
<summary>Requires successful base and owned Assertion initialization.</summary>
*)
{endregion}
METHOD PROTECTED CheckInitialization : BOOL //! TRUE when the inherited initialization check and this concrete fixture check both accept the setup.
CheckInitialization := FALSE;
IF NOT SUPER^.CheckInitialization() THEN
    RETURN;
END_IF;

CheckInitialization := FDuplicateRejected.IsInitialized
    AND FNullRejected.IsInitialized
    AND FExplicitSlotRejected.IsInitialized
    AND FMissingSlotRejected.IsInitialized
    AND FZeroSlotRejected.IsInitialized
    AND FSlotGapRejected.IsInitialized;
END_METHOD

{region 'Documentation'}
(*!
<summary>Configures one direct builder scenario and its named Assertions.</summary>
*)
{endregion}
METHOD PROTECTED Configure
FPreparationStateCount := 0;
FTestStateCount := 1;
FScenarioExecuted := FALSE;
FChecksEvaluated := FALSE;

FDuplicateRejectedMatches := FALSE;
FDuplicateRejected.Initialize(Parent := THIS^,
    AssertionName := 'DuplicateRejected');
FNullRejectedMatches := FALSE;
FNullRejected.Initialize(Parent := THIS^,
    AssertionName := 'NullRejected');
FExplicitSlotRejectedMatches := FALSE;
FExplicitSlotRejected.Initialize(Parent := THIS^,
    AssertionName := 'ExplicitSlotRejected');
FMissingSlotRejectedMatches := FALSE;
FMissingSlotRejected.Initialize(Parent := THIS^,
    AssertionName := 'MissingSlotRejected');
FZeroSlotRejectedMatches := FALSE;
FZeroSlotRejected.Initialize(Parent := THIS^,
    AssertionName := 'ZeroSlotRejected');
FSlotGapRejectedMatches := FALSE;
FSlotGapRejected.Initialize(Parent := THIS^,
    AssertionName := 'SlotGapRejected');
END_METHOD

{region 'Documentation'}
(*!
<summary>Completes Abort immediately; no asynchronous resource operation is started.</summary>
*)
{endregion}
METHOD PROTECTED ProcessAbort
VAR_INPUT
    Enable : BOOL; //! Phase permission supplied by the owning Test Case; FALSE does not authorize progression, while observation may continue.
END_VAR
IF Enable THEN
    CompleteAbort();
END_IF;
END_METHOD

{region 'Documentation'}
(*!
<summary>Evaluates recorded observations and consumes pending resets on disabled calls.</summary>
*)
{endregion}
METHOD PROTECTED ProcessAssertions
VAR_INPUT
    Enable : BOOL; //! Phase permission supplied by the owning Test Case; FALSE does not authorize progression, while observation may continue.
END_VAR
FDuplicateRejected(Enable := Enable,
    State := State,
    IN := FDuplicateRejectedMatches);

FNullRejected(Enable := Enable,
    State := State,
    IN := FNullRejectedMatches);

FExplicitSlotRejected(Enable := Enable,
    State := State,
    IN := FExplicitSlotRejectedMatches);

FMissingSlotRejected(Enable := Enable,
    State := State,
    IN := FMissingSlotRejectedMatches);

FZeroSlotRejected(Enable := Enable,
    State := State,
    IN := FZeroSlotRejectedMatches);

FSlotGapRejected(Enable := Enable,
    State := State,
    IN := FSlotGapRejectedMatches);

IF Enable AND FDuplicateRejected.EvaluationActive
    AND FNullRejected.EvaluationActive
    AND FExplicitSlotRejected.EvaluationActive
    AND FMissingSlotRejected.EvaluationActive
    AND FZeroSlotRejected.EvaluationActive
    AND FSlotGapRejected.EvaluationActive THEN
    FChecksEvaluated := TRUE;
END_IF;
END_METHOD

{region 'Documentation'}
(*!
<summary>No Preparation phase is needed for synchronous builder calls.</summary>
*)
{endregion}
METHOD PROTECTED ProcessPreparations
VAR_INPUT
    // SA0033: Required override signature; this scenario has no Preparation work.
    {attribute 'analysis' := '-33'}
    Enable : BOOL; //! Phase permission supplied by the owning Test Case; FALSE does not authorize progression, while observation may continue.
END_VAR
END_METHOD

{region 'Documentation'}
(*!
<summary>Clears recorded checks and Assertion results; each scenario initializes its own builder.</summary>
*)
{endregion}
METHOD PROTECTED ProcessReset
FScenarioExecuted := FALSE;
FChecksEvaluated := FALSE;
FDuplicateRejectedMatches := FALSE;
FDuplicateRejected.Reset();
FNullRejectedMatches := FALSE;
FNullRejected.Reset();
FExplicitSlotRejectedMatches := FALSE;
FExplicitSlotRejected.Reset();
FMissingSlotRejectedMatches := FALSE;
FMissingSlotRejected.Reset();
FZeroSlotRejectedMatches := FALSE;
FZeroSlotRejected.Reset();
FSlotGapRejectedMatches := FALSE;
FSlotGapRejected.Reset();
CompleteReset();
END_METHOD

{region 'Documentation'}
(*!
<summary>Runs setup operations once, then completes after their observations have been evaluated.</summary>
*)
{endregion}
METHOD PROTECTED ProcessTests
VAR_INPUT
    Enable : BOOL; //! Phase permission supplied by the owning Test Case; FALSE does not authorize progression, while observation may continue.
END_VAR
IF NOT Enable THEN
    RETURN;
END_IF;

IF FChecksEvaluated THEN
    CompleteTests();
ELSIF NOT FScenarioExecuted THEN
    RunScenario();
    FScenarioExecuted := TRUE;
END_IF;
END_METHOD

{region 'Documentation'}
(*!
<summary>Checks typical setup mistakes without executing the registered child objects.</summary>
*)
{endregion}
METHOD PRIVATE RunScenario
VAR
    ChildA : I_TestSuite;
    ChildB : I_TestSuite;
    AcceptedA : BOOL;
    AcceptedB : BOOL;
    Config : ST_TestSuiteCollectionConfig;
    AcceptedAfterError : BOOL;
END_VAR
ChildA := FChildA;
ChildB := FChildB;
FBuilder.Initialize(Mode := E_OrchestrationMode.Serial,
    TestSuites := FSuites);
AcceptedA := FBuilder.Register(TestSuite := ChildA);
AcceptedB := FBuilder.Register(TestSuite := ChildA);
AcceptedAfterError := FBuilder.Register(TestSuite := ChildB);
Config := FBuilder.Finalize();
FDuplicateRejectedMatches := AcceptedA AND NOT AcceptedB AND NOT AcceptedAfterError
    AND NOT Config.IsValid AND (FBuilder.Count = 1)
    AND (FSuites[1] = ChildA) AND (FSuites[2] = 0) AND (FChildA.ExecutionSlot = 1);

FBuilder.Initialize(Mode := E_OrchestrationMode.Serial,
    TestSuites := FSuites);
AcceptedA := FBuilder.Register(TestSuite := ChildA);
AcceptedB := FBuilder.Register(TestSuite := 0);
Config := FBuilder.Finalize();
FNullRejectedMatches := AcceptedA AND NOT AcceptedB AND NOT Config.IsValid
    AND (FBuilder.Count = 1) AND (FSuites[1] = ChildA) AND (FSuites[2] = 0);

FBuilder.Initialize(Mode := E_OrchestrationMode.Serial,
    TestSuites := FSuites);
FChildA.ExecutionSlot := CandidateSlotBeforeRejection;
AcceptedA := FBuilder.RegisterWithSlot(TestSuite := ChildA,
    ExecutionSlot := 1);
Config := FBuilder.Finalize();
FExplicitSlotRejectedMatches := NOT AcceptedA AND NOT Config.IsValid
    AND (FBuilder.Count = 0) AND (FSuites[1] = 0)
    AND (FChildA.ExecutionSlot = CandidateSlotBeforeRejection);

FBuilder.Initialize(Mode := E_OrchestrationMode.ParallelSlots,
    TestSuites := FSuites);
AcceptedA := FBuilder.Register(TestSuite := ChildA);
Config := FBuilder.Finalize();
FMissingSlotRejectedMatches := NOT AcceptedA AND NOT Config.IsValid
    AND (FBuilder.Count = 0) AND (FSuites[1] = 0)
    AND (FChildA.ExecutionSlot = CandidateSlotBeforeRejection);

FBuilder.Initialize(Mode := E_OrchestrationMode.ParallelSlots,
    TestSuites := FSuites);
AcceptedA := FBuilder.RegisterWithSlot(TestSuite := ChildA,
    ExecutionSlot := 0);
Config := FBuilder.Finalize();
FZeroSlotRejectedMatches := NOT AcceptedA AND NOT Config.IsValid
    AND (FBuilder.Count = 0) AND (FSuites[1] = 0)
    AND (FChildA.ExecutionSlot = CandidateSlotBeforeRejection);

FBuilder.Initialize(Mode := E_OrchestrationMode.ParallelSlots,
    TestSuites := FSuites);
AcceptedA := FBuilder.RegisterWithSlot(TestSuite := ChildA,
    ExecutionSlot := 1);
AcceptedB := FBuilder.RegisterWithSlot(TestSuite := ChildB,
    ExecutionSlot := 3);
Config := FBuilder.Finalize();
FSlotGapRejectedMatches := AcceptedA AND AcceptedB AND NOT Config.IsValid
    AND FBuilder.IsFinalized AND (FBuilder.Count = 2)
    AND (FSuites[1] = ChildA) AND (FSuites[2] = ChildB);
END_METHOD

END_FUNCTION_BLOCK

// ---- SelfTests/TestCases/TestSuite_RunControlConfigurationBuilder/Test_RunControlBuilderFinalizeReuse.TcPOU
{region 'Documentation'}
(*!
<summary>Checks empty and repeated finalization, sealed registration and a clean new build.</summary>
<description>Child mocks are inert interface identities and slot storage only; no child initialization or FB call is performed.</description>
*)
{endregion}
FUNCTION_BLOCK Test_RunControlBuilderFinalizeReuse EXTENDS TestCaseBase
VAR
    FBuilder : RunControlConfigurationBuilder;
    FSuites : ARRAY[1..2] OF I_TestSuite;
    FChildA : TestSuiteMock;
    FChildB : TestSuiteMock;
    FScenarioExecuted : BOOL;
    FChecksEvaluated : BOOL;
    FEmptyRejected : AssertTrue;
    FEmptyRejectedMatches : BOOL;
    FRepeatedFinalization : AssertTrue;
    FRepeatedFinalizationMatches : BOOL;
    FSealedRegistration : AssertTrue;
    FSealedRegistrationMatches : BOOL;
    FErrorRecorded : AssertTrue;
    FErrorRecordedMatches : BOOL;
    FFreshInitialize : AssertTrue;
    FFreshInitializeMatches : BOOL;
    FReuse : AssertTrue;
    FReuseMatches : BOOL;
END_VAR
VAR CONSTANT
    CandidateSlotBeforeRejection : UINT := 9;
END_VAR

SUPER^();

{region 'Documentation'}
(*!
<summary>Contributes each owned Assertion once without executing it.</summary>
*)
{endregion}
METHOD PROTECTED AggregateResults
VAR_INPUT
    Aggregator : I_ResultAggregator; //! Borrowed result sink owned by the outer Test Case; add this test's checking Assertions without resetting or retaining the sink.
END_VAR
Aggregator.AddProvider(Provider := FEmptyRejected);
Aggregator.AddProvider(Provider := FRepeatedFinalization);
Aggregator.AddProvider(Provider := FSealedRegistration);
Aggregator.AddProvider(Provider := FErrorRecorded);
Aggregator.AddProvider(Provider := FFreshInitialize);
Aggregator.AddProvider(Provider := FReuse);
END_METHOD

{region 'Documentation'}
(*!
<summary>Requires successful base and owned Assertion initialization.</summary>
*)
{endregion}
METHOD PROTECTED CheckInitialization : BOOL //! TRUE when the inherited initialization check and this concrete fixture check both accept the setup.
CheckInitialization := FALSE;
IF NOT SUPER^.CheckInitialization() THEN
    RETURN;
END_IF;

CheckInitialization := FEmptyRejected.IsInitialized
    AND FRepeatedFinalization.IsInitialized
    AND FSealedRegistration.IsInitialized
    AND FErrorRecorded.IsInitialized
    AND FFreshInitialize.IsInitialized
    AND FReuse.IsInitialized;
END_METHOD

{region 'Documentation'}
(*!
<summary>Configures one direct builder scenario and its named Assertions.</summary>
*)
{endregion}
METHOD PROTECTED Configure
FPreparationStateCount := 0;
FTestStateCount := 1;
FScenarioExecuted := FALSE;
FChecksEvaluated := FALSE;

FEmptyRejectedMatches := FALSE;
FEmptyRejected.Initialize(Parent := THIS^,
    AssertionName := 'EmptyRejected');
FRepeatedFinalizationMatches := FALSE;
FRepeatedFinalization.Initialize(Parent := THIS^,
    AssertionName := 'RepeatedFinalization');
FSealedRegistrationMatches := FALSE;
FSealedRegistration.Initialize(Parent := THIS^,
    AssertionName := 'SealedRegistration');
FErrorRecordedMatches := FALSE;
FErrorRecorded.Initialize(Parent := THIS^,
    AssertionName := 'ErrorRecorded');
FFreshInitializeMatches := FALSE;
FFreshInitialize.Initialize(Parent := THIS^,
    AssertionName := 'FreshInitialize');
FReuseMatches := FALSE;
FReuse.Initialize(Parent := THIS^,
    AssertionName := 'Reuse');
END_METHOD

{region 'Documentation'}
(*!
<summary>Completes Abort immediately; no asynchronous resource operation is started.</summary>
*)
{endregion}
METHOD PROTECTED ProcessAbort
VAR_INPUT
    Enable : BOOL; //! Phase permission supplied by the owning Test Case; FALSE does not authorize progression, while observation may continue.
END_VAR
IF Enable THEN
    CompleteAbort();
END_IF;
END_METHOD

{region 'Documentation'}
(*!
<summary>Evaluates recorded observations and consumes pending resets on disabled calls.</summary>
*)
{endregion}
METHOD PROTECTED ProcessAssertions
VAR_INPUT
    Enable : BOOL; //! Phase permission supplied by the owning Test Case; FALSE does not authorize progression, while observation may continue.
END_VAR
FEmptyRejected(Enable := Enable,
    State := State,
    IN := FEmptyRejectedMatches);

FRepeatedFinalization(Enable := Enable,
    State := State,
    IN := FRepeatedFinalizationMatches);

FSealedRegistration(Enable := Enable,
    State := State,
    IN := FSealedRegistrationMatches);

FErrorRecorded(Enable := Enable,
    State := State,
    IN := FErrorRecordedMatches);

FFreshInitialize(Enable := Enable,
    State := State,
    IN := FFreshInitializeMatches);

FReuse(Enable := Enable,
    State := State,
    IN := FReuseMatches);

IF Enable AND FEmptyRejected.EvaluationActive
    AND FRepeatedFinalization.EvaluationActive
    AND FSealedRegistration.EvaluationActive
    AND FErrorRecorded.EvaluationActive
    AND FFreshInitialize.EvaluationActive
    AND FReuse.EvaluationActive THEN
    FChecksEvaluated := TRUE;
END_IF;
END_METHOD

{region 'Documentation'}
(*!
<summary>No Preparation phase is needed for synchronous builder calls.</summary>
*)
{endregion}
METHOD PROTECTED ProcessPreparations
VAR_INPUT
    // SA0033: Required override signature; this scenario has no Preparation work.
    {attribute 'analysis' := '-33'}
    Enable : BOOL; //! Phase permission supplied by the owning Test Case; FALSE does not authorize progression, while observation may continue.
END_VAR
END_METHOD

{region 'Documentation'}
(*!
<summary>Clears recorded checks and Assertion results; each scenario initializes its own builder.</summary>
*)
{endregion}
METHOD PROTECTED ProcessReset
FScenarioExecuted := FALSE;
FChecksEvaluated := FALSE;
FEmptyRejectedMatches := FALSE;
FEmptyRejected.Reset();
FRepeatedFinalizationMatches := FALSE;
FRepeatedFinalization.Reset();
FSealedRegistrationMatches := FALSE;
FSealedRegistration.Reset();
FErrorRecordedMatches := FALSE;
FErrorRecorded.Reset();
FFreshInitializeMatches := FALSE;
FFreshInitialize.Reset();
FReuseMatches := FALSE;
FReuse.Reset();
CompleteReset();
END_METHOD

{region 'Documentation'}
(*!
<summary>Runs setup operations once, then completes after their observations have been evaluated.</summary>
*)
{endregion}
METHOD PROTECTED ProcessTests
VAR_INPUT
    Enable : BOOL; //! Phase permission supplied by the owning Test Case; FALSE does not authorize progression, while observation may continue.
END_VAR
IF NOT Enable THEN
    RETURN;
END_IF;

IF FChecksEvaluated THEN
    CompleteTests();
ELSIF NOT FScenarioExecuted THEN
    RunScenario();
    FScenarioExecuted := TRUE;
END_IF;
END_METHOD

{region 'Documentation'}
(*!
<summary>Checks empty and repeated finalization, sealed registration and a clean new build.</summary>
*)
{endregion}
METHOD PRIVATE RunScenario
VAR
    ChildA : I_TestSuite;
    ChildB : I_TestSuite;
    AcceptedA : BOOL;
    AcceptedB : BOOL;
    Config : ST_TestSuiteCollectionConfig;
    RepeatedConfig : ST_TestSuiteCollectionConfig;
END_VAR
ChildA := FChildA;
ChildB := FChildB;
FBuilder.Initialize(Mode := E_OrchestrationMode.Serial,
    TestSuites := FSuites);
Config := FBuilder.Finalize();
RepeatedConfig := FBuilder.Finalize();
FEmptyRejectedMatches := NOT Config.IsValid AND NOT RepeatedConfig.IsValid
    AND FBuilder.IsFinalized AND NOT FBuilder.IsValid AND (RepeatedConfig.Count = 0);

FBuilder.Initialize(Mode := E_OrchestrationMode.Serial,
    TestSuites := FSuites);
AcceptedA := FBuilder.Register(TestSuite := ChildA);
Config := FBuilder.Finalize();
RepeatedConfig := FBuilder.Finalize();
FRepeatedFinalizationMatches := AcceptedA AND Config.IsValid AND RepeatedConfig.IsValid
    AND (RepeatedConfig.FirstIndex = Config.FirstIndex)
    AND (RepeatedConfig.LastIndex = Config.LastIndex)
    AND (RepeatedConfig.Count = Config.Count) AND (RepeatedConfig.Mode = Config.Mode);

FChildB.ExecutionSlot := CandidateSlotBeforeRejection;
AcceptedB := FBuilder.Register(TestSuite := ChildB);
RepeatedConfig := FBuilder.Finalize();
FSealedRegistrationMatches := NOT AcceptedB AND RepeatedConfig.IsValid AND FBuilder.IsValid
    AND FBuilder.IsFinalized AND (FBuilder.Count = 1)
    AND (FSuites[1] = ChildA) AND (FSuites[2] = 0)
    AND (FChildB.ExecutionSlot = CandidateSlotBeforeRejection);

FBuilder.Initialize(Mode := E_OrchestrationMode.Serial,
    TestSuites := FSuites);
AcceptedA := FBuilder.Register(TestSuite := ChildA);
AcceptedB := FBuilder.Register(TestSuite := ChildA);
Config := FBuilder.Finalize();
FErrorRecordedMatches := AcceptedA AND NOT AcceptedB AND NOT Config.IsValid;

FBuilder.Initialize(Mode := E_OrchestrationMode.Parallel,
    TestSuites := FSuites);
FFreshInitializeMatches := NOT FBuilder.IsFinalized AND NOT FBuilder.IsValid
    AND (FBuilder.Count = 0) AND (FBuilder.Mode = E_OrchestrationMode.Parallel)
    AND (FSuites[1] = 0) AND (FSuites[2] = 0);
AcceptedB := FBuilder.Register(TestSuite := ChildB);
Config := FBuilder.Finalize();
FReuseMatches := AcceptedB AND Config.IsValid AND FBuilder.IsValid AND FBuilder.IsFinalized
    AND (Config.Count = 1) AND (Config.Mode = E_OrchestrationMode.Parallel)
    AND (FSuites[1] = ChildB) AND (FSuites[2] = 0) AND (FChildB.ExecutionSlot = 1);
END_METHOD

END_FUNCTION_BLOCK

// ---- SelfTests/TestSuites/TestSuite_TestSuiteLifecycle.TcPOU
{region 'Documentation'}
(*!
<summary>Groups isolated Suite owner tests; detailed scheduling remains in its own suites.</summary>
*)
{endregion}
FUNCTION_BLOCK TestSuite_TestSuiteLifecycle EXTENDS TestSuiteBase
VAR
    FSubjectParent : I_RunControl;
    FInitialization : Test_SuiteInitialization;
    FReadiness : Test_SuiteReadiness;
    FNormalCompletion : Test_SuiteNormalLifecycle;
    FMixedResults : Test_SuiteNormalLifecycle;
    FTestCases : ARRAY[1..TestCaseCapacity] OF I_TestCase;
    FResetError : Test_SuiteExceptionalLifecycle;
    FResetTimeout : Test_SuiteExceptionalLifecycle;
    FChildError : Test_SuiteExceptionalLifecycle;
    FUnexpectedChildAbort : Test_SuiteExceptionalLifecycle;
    FExecutionError : Test_SuiteExceptionalLifecycle;
    FExecutionTimeout : Test_SuiteExceptionalLifecycle;
    FAbort : Test_SuiteExceptionalLifecycle;
    FAbortError : Test_SuiteExceptionalLifecycle;
    FAbortTimeout : Test_SuiteExceptionalLifecycle;
    FFinalization : Test_SuiteFinalization;
    FLateResetChildren : Test_SuiteFinalization;
    FReservationRelease : Test_SuiteReservationRelease;
    FRealComposition : Test_SuiteRealComposition;
    FMockRepeatedReset : Test_SuiteMockRepeatedReset;
END_VAR
VAR CONSTANT
    TestCaseCapacity : UINT := 18;
END_VAR

SUPER^();

{region 'Documentation'}
(*!
<summary>Supplies the existing root identity for isolated Suite subjects before this Suite is initialized.</summary>
*)
{endregion}
METHOD PUBLIC BindSubjectParent
VAR_INPUT
    Parent : I_RunControl; //! Borrowed identity parent retained for isolated subject initialization; keep the Run-Control alive through subject use.
END_VAR
FSubjectParent := Parent;
END_METHOD

{region 'Documentation'}
(*!
<summary>Initializes and registers independent Suite-owner scenarios for serial execution.</summary>
*)
{endregion}
METHOD PROTECTED Configure
VAR_IN_OUT
    // SA0167: Borrowed owner builder; no temporary instance is created.
    {attribute 'analysis' := '-167'}
    Builder : TestSuiteConfigurationBuilder; //! Borrowed owner configuration builder used only during this Configure call; register this owner's concrete children.
END_VAR
VAR
    TestConfig : ST_TestCaseConfig;
END_VAR
Builder.Initialize(Mode := E_OrchestrationMode.Serial,
    TestCases := FTestCases);
FInitialization.BindSubjectParent(Parent := FSubjectParent);
FInitialization.Initialize(Parent := THIS^,
    TestName := 'Initialization',
    Config := TestConfig);
Builder.Register(TestCase := FInitialization);
FReadiness.BindSubjectParent(Parent := FSubjectParent);
FReadiness.Initialize(Parent := THIS^,
    TestName := 'Readiness',
    Config := TestConfig);
Builder.Register(TestCase := FReadiness);

FNormalCompletion.BindSubjectParent(Parent := FSubjectParent);
FNormalCompletion.Initialize(Parent := THIS^,
    TestName := 'NormalCompletion',
    Config := TestConfig);
Builder.Register(TestCase := FNormalCompletion);

FMixedResults.BindSubjectParent(Parent := FSubjectParent);
FMixedResults.Initialize(Parent := THIS^,
    TestName := 'MixedResults',
    Config := TestConfig);
Builder.Register(TestCase := FMixedResults);

FResetError.BindSubjectParent(Parent := FSubjectParent);
FResetError.Initialize(Parent := THIS^,
    TestName := 'ResetError',
    Config := TestConfig);
Builder.Register(TestCase := FResetError);

FResetTimeout.BindSubjectParent(Parent := FSubjectParent);
FResetTimeout.Initialize(Parent := THIS^,
    TestName := 'ResetTimeout',
    Config := TestConfig);
Builder.Register(TestCase := FResetTimeout);

FChildError.BindSubjectParent(Parent := FSubjectParent);
FChildError.Initialize(Parent := THIS^,
    TestName := 'ChildError',
    Config := TestConfig);
Builder.Register(TestCase := FChildError);

FUnexpectedChildAbort.BindSubjectParent(Parent := FSubjectParent);
FUnexpectedChildAbort.Initialize(Parent := THIS^,
    TestName := 'UnexpectedChildAbort',
    Config := TestConfig);
Builder.Register(TestCase := FUnexpectedChildAbort);

FExecutionError.BindSubjectParent(Parent := FSubjectParent);
FExecutionError.Initialize(Parent := THIS^,
    TestName := 'ExecutionError',
    Config := TestConfig);
Builder.Register(TestCase := FExecutionError);

FExecutionTimeout.BindSubjectParent(Parent := FSubjectParent);
FExecutionTimeout.Initialize(Parent := THIS^,
    TestName := 'ExecutionTimeout',
    Config := TestConfig);
Builder.Register(TestCase := FExecutionTimeout);

FAbort.BindSubjectParent(Parent := FSubjectParent);
FAbort.Initialize(Parent := THIS^,
    TestName := 'Abort',
    Config := TestConfig);
Builder.Register(TestCase := FAbort);

FAbortError.BindSubjectParent(Parent := FSubjectParent);
FAbortError.Initialize(Parent := THIS^,
    TestName := 'AbortError',
    Config := TestConfig);
Builder.Register(TestCase := FAbortError);

FAbortTimeout.BindSubjectParent(Parent := FSubjectParent);
FAbortTimeout.Initialize(Parent := THIS^,
    TestName := 'AbortTimeout',
    Config := TestConfig);
Builder.Register(TestCase := FAbortTimeout);

FFinalization.BindSubjectParent(Parent := FSubjectParent);
FFinalization.Initialize(Parent := THIS^,
    TestName := 'Finalization',
    Config := TestConfig);
Builder.Register(TestCase := FFinalization);

FLateResetChildren.BindSubjectParent(Parent := FSubjectParent);
FLateResetChildren.Initialize(Parent := THIS^,
    TestName := 'LateResetChildren',
    Config := TestConfig);
Builder.Register(TestCase := FLateResetChildren);

FReservationRelease.BindSubjectParent(Parent := FSubjectParent);
FReservationRelease.Initialize(Parent := THIS^,
    TestName := 'ReservationRelease',
    Config := TestConfig);
Builder.Register(TestCase := FReservationRelease);

FRealComposition.BindSubjectParent(Parent := FSubjectParent);
FRealComposition.Initialize(Parent := THIS^,
    TestName := 'RealComposition',
    Config := TestConfig);
Builder.Register(TestCase := FRealComposition);

FMockRepeatedReset.BindSubjectParent(Parent := FSubjectParent);
FMockRepeatedReset.Initialize(Parent := THIS^,
    TestName := 'MockRepeatedReset',
    Config := TestConfig);
Builder.Register(TestCase := FMockRepeatedReset);
END_METHOD

{region 'Documentation'}
(*!
<summary>Returns a registered scenario using its original array index.</summary>
*)
{endregion}
METHOD PUBLIC GetTestCase : I_TestCase //! Typed child interface at the original array index; zero when no entry is available.
VAR_INPUT
    Index : DINT; //! Original occupied child-array index, rather than an ordinal position.
END_VAR
GetTestCase := 0;
IF (ChildCount = 0) OR (Index < ChildArrayLowerBound)
    OR (DINT_TO_LINT(Index) >= DINT_TO_LINT(ChildArrayLowerBound) + UINT_TO_LINT(ChildCount)) THEN
    RETURN;
END_IF;
GetTestCase := FTestCases[Index];
END_METHOD

{region 'Documentation'}
(*!
<summary>Calls each owned scenario once per initialized Suite cycle.</summary>
*)
{endregion}
METHOD PROTECTED ProcessTestCases
FInitialization();
FReadiness();
FNormalCompletion(FirstChildResult := E_Result.Passed);
FMixedResults(FirstChildResult := E_Result.Failed);

FResetError(Scenario := E_SuiteLifecycleScenario.ResetError);
FResetTimeout(Scenario := E_SuiteLifecycleScenario.ResetTimeout);
FChildError(Scenario := E_SuiteLifecycleScenario.ChildError);
FUnexpectedChildAbort(Scenario := E_SuiteLifecycleScenario.UnexpectedChildAbort);
FExecutionError(Scenario := E_SuiteLifecycleScenario.ExecutionError);
FExecutionTimeout(Scenario := E_SuiteLifecycleScenario.ExecutionTimeout);
FAbort(Scenario := E_SuiteLifecycleScenario.Abort);
FAbortError(Scenario := E_SuiteLifecycleScenario.AbortError);
FAbortTimeout(Scenario := E_SuiteLifecycleScenario.AbortTimeout);

FFinalization(LateResetChildren := FALSE);
FLateResetChildren(LateResetChildren := TRUE);
FReservationRelease();

FRealComposition();
FMockRepeatedReset();
END_METHOD

END_FUNCTION_BLOCK

// ---- SelfTests/TestCases/TestSuite_TestSuiteLifecycle/Test_SuiteInitialization.TcPOU
{region 'Documentation'}
(*!
<summary>Checks Suite initialization, collection handover, rejected setup and passivity before parent Reset.</summary>
<description>
Each Test state is one setup attempt, followed by two subject calls without lifecycle requests.
Valid setup comes first and last: intervening rejected attempts must not reuse a previously
valid collection. This represents successive startup configurations, not hot reconfiguration.
Identity failures precede Configure; builder failure precedes helper initialization; later
configuration failures hide the collection again. The helper queries it during Initialize.
The subject and its initialization diagnostics use the local capture. Checking Assertions
use the outer selftest publisher and retain failures across all attempts.
</description>
*)
{endregion}
FUNCTION_BLOCK Test_SuiteInitialization EXTENDS TestCaseBase
VAR
    FSubjectParent : I_RunControl;
    FSubject : TestSuiteLifecycleProbe;
    FHelper : SuiteOrchestratorDouble;
    FCapture : EventBuffer;
    FEvents : ARRAY[1..CaptureLength] OF ST_Event;
    FCaptureFifo : ST_FifoStatus;
    FCaptureStatus : ST_EventBufferStatus;
    FFixtureValid : BOOL;
    FAttempt : INT := FirstValidSetup;
    FAttemptStarted : BOOL;
    FChecked : BOOL;
    FPassiveCalls : UINT;
    FExpectedInitialized : BOOL;
    FInitialSequence : UDINT;
    FInitialization : AssertTrue;
    FInitializationMatches : BOOL;
    FConfigureOrder : AssertTrue;
    FConfigureOrderMatches : BOOL;
    FCollection : AssertTrue;
    FCollectionMatches : BOOL;
    FPassiveState : AssertTrue;
    FPassiveStateMatches : BOOL;
    FDiagnostic : AssertTrue;
    FDiagnosticMatches : BOOL;
    FDispatch : AssertTrue;
    FDispatchMatches : BOOL;
    FCaptureIntegrity : AssertTrue;
END_VAR
VAR CONSTANT
    CaptureLength : UINT := 32;
    PassiveCallCount : UINT := 2;
    FirstValidSetup : INT := 1;
    MissingParent : INT := 2;
    InvalidName : INT := 3;
    OverlengthName : INT := 4;
    NoRegistration : INT := 5;
    UninitializedChild : INT := 6;
    ZeroExecutionTimeout : INT := 7;
    ZeroResetTimeout : INT := 8;
    ZeroAbortTimeout : INT := 9;
    RejectedHelper : INT := 10;
    FinalValidSetup : INT := 11;
    AttemptCount : INT := 11;
END_VAR

SUPER^();

